(* IEC 61131-3 sources: daoli-st-library/DL_MathData (part 10) *)

(* ---- FC_DL_CharIsAlnum.st ---- *)
(*==============================================================================
 * 组件名称 : FC_DL_CharIsAlnum ｜ 子库 : DL_MathData ｜ v1.0.0 ｜ 2026-11-23
 * 平台     : CODESYS 3.5 / TwinCAT 3 / InoProShop / Machine Expert（纯 IEC，无厂商库）
 * 功能简介 : 判定 STRING(1) 单字符是否为字母或数字（'0'..'9' / 'A'..'Z' /
 *            'a'..'z'），直接以字符（ASCII 序）比较实现，不用库函数。
 * 契约     : 返回 TRUE = 字母或数字；输入 sChar 单字符，空串恒 FALSE；
 *            纯函数无状态、同输入同输出。
 * 开源溯源 : 来源 fisothemes/TwinCAT-Dynamic-String-Kit
 *            https://github.com/fisothemes/TwinCAT-Dynamic-String-Kit / MIT
 *            借鉴点：字符分类谓词语义，实现为本库 clean-room 重写。
 * 依赖     : 无 DL_ 内部依赖（本批自足实现）
 * 红线自检 : R1 零全局 R2 零%I/%Q R3 纯IEC R4 空串防御（区间外恒 FALSE）
 *            R5 双语注释 R6 N/A（无状态机） R7 N/A（无定时器实例）
 * 修订历史 : 2026-11-23 R78-B1 字符分类族模板派生首版
 *============================================================================*)
FUNCTION FC_DL_CharIsAlnum : BOOL
VAR_INPUT
    sChar : STRING(1);      // 待判定单字符（空串恒 FALSE） / Single character to test (empty = FALSE)
END_VAR
IF (sChar >= '0') AND (sChar <= '9') THEN
    FC_DL_CharIsAlnum := TRUE;      // 数字字符命中 / Digit hit
ELSIF ((sChar >= 'A') AND (sChar <= 'Z')) OR ((sChar >= 'a') AND (sChar <= 'z')) THEN
    FC_DL_CharIsAlnum := TRUE;      // 字母字符命中 / Letter hit
ELSE
    FC_DL_CharIsAlnum := FALSE;     // 空串或其他字符 / Empty string or other character
END_IF
END_FUNCTION

(* ---- FC_DL_CharIsAlpha.st ---- *)
(*==============================================================================
 * 组件名称 : FC_DL_CharIsAlpha ｜ 子库 : DL_MathData ｜ v1.0.0 ｜ 2026-11-23
 * 平台     : CODESYS 3.5 / TwinCAT 3 / InoProShop / Machine Expert（纯 IEC，无厂商库）
 * 功能简介 : 判定 STRING(1) 单字符是否为英文字母 'A'..'Z' 或 'a'..'z'，
 *            直接以字符（ASCII 序）比较实现，不调用任何字符分类库函数。
 * 契约     : 返回 TRUE = 英文字母；输入 sChar 单字符，空串按非字母处理；
 *            纯函数无状态、同输入同输出。
 * 开源溯源 : 来源 fisothemes/TwinCAT-Dynamic-String-Kit
 *            https://github.com/fisothemes/TwinCAT-Dynamic-String-Kit / MIT
 *            借鉴点：字符分类谓词语义，实现为本库 clean-room 重写。
 * 依赖     : 无 DL_ 内部依赖（本批自足实现）
 * 红线自检 : R1 零全局 R2 零%I/%Q R3 纯IEC R4 空串防御（区间外恒 FALSE）
 *            R5 双语注释 R6 N/A（无状态机） R7 N/A（无定时器实例）
 * 修订历史 : 2026-11-23 R78-B1 字符分类族模板派生首版
 *============================================================================*)
FUNCTION FC_DL_CharIsAlpha : BOOL
VAR_INPUT
    sChar : STRING(1);      // 待判定单字符（空串按非字母） / Single character to test (empty = not alpha)
END_VAR
IF ((sChar >= 'A') AND (sChar <= 'Z')) OR ((sChar >= 'a') AND (sChar <= 'z')) THEN
    FC_DL_CharIsAlpha := TRUE;      // 命中大小写字母区间 / Within letter ranges A-Z or a-z
ELSE
    FC_DL_CharIsAlpha := FALSE;     // 空串或非字母字符 / Empty string or non-letter
END_IF
END_FUNCTION

(* ---- FC_DL_CharIsDigit.st ---- *)
(*==============================================================================
 * 组件名称 : FC_DL_CharIsDigit ｜ 子库 : DL_MathData ｜ v1.0.0 ｜ 2026-11-23
 * 平台     : CODESYS 3.5 / TwinCAT 3 / InoProShop / Machine Expert（纯 IEC，无厂商库）
 * 功能简介 : 判定 STRING(1) 单字符是否为十进制数字字符 '0'..'9'，
 *            直接以字符（ASCII 序）比较实现，不调用任何字符分类库函数。
 * 契约     : 返回 TRUE = 数字字符；输入 sChar 单字符，空串按非数字处理；
 *            纯函数无状态、同输入同输出。
 * 开源溯源 : 来源 fisothemes/TwinCAT-Dynamic-String-Kit
 *            https://github.com/fisothemes/TwinCAT-Dynamic-String-Kit / MIT
 *            借鉴点：字符分类谓词语义，实现为本库 clean-room 重写。
 * 依赖     : 无 DL_ 内部依赖（本批自足实现）
 * 红线自检 : R1 零全局 R2 零%I/%Q R3 纯IEC R4 空串防御（区间外恒 FALSE）
 *            R5 双语注释 R6 N/A（无状态机） R7 N/A（无定时器实例）
 * 修订历史 : 2026-11-23 R78-B1 字符分类族模板派生首版
 *============================================================================*)
FUNCTION FC_DL_CharIsDigit : BOOL
VAR_INPUT
    sChar : STRING(1);      // 待判定单字符（空串按非数字） / Single character to test (empty = not a digit)
END_VAR
IF (sChar >= '0') AND (sChar <= '9') THEN
    FC_DL_CharIsDigit := TRUE;      // 命中 '0'..'9' 区间 / Within digit range '0'..'9'
ELSE
    FC_DL_CharIsDigit := FALSE;     // 空串或非数字字符 / Empty string or non-digit
END_IF
END_FUNCTION

(* ---- FC_DL_CharIsHexDigit.st ---- *)
(*==============================================================================
 * 组件名称 : FC_DL_CharIsHexDigit ｜ 子库 : DL_MathData ｜ v1.0.0 ｜ 2026-11-23
 * 平台     : CODESYS 3.5 / TwinCAT 3 / InoProShop / Machine Expert（纯 IEC，无厂商库）
 * 功能简介 : 判定 STRING(1) 单字符是否为十六进制位（'0'..'9' / 'A'..'F' /
 *            'a'..'f'），直接以字符（ASCII 序）比较实现，不用库函数。
 * 契约     : 返回 TRUE = 十六进制位；输入 sChar 单字符，空串恒 FALSE；
 *            纯函数无状态、同输入同输出。
 * 开源溯源 : 来源 fisothemes/TwinCAT-Dynamic-String-Kit
 *            https://github.com/fisothemes/TwinCAT-Dynamic-String-Kit / MIT
 *            借鉴点：字符分类谓词语义，实现为本库 clean-room 重写。
 * 依赖     : 无 DL_ 内部依赖（本批自足实现）
 * 红线自检 : R1 零全局 R2 零%I/%Q R3 纯IEC R4 空串防御（恒 FALSE）
 *            R5 双语注释 R6 N/A（无状态机） R7 N/A（无定时器实例）
 * 修订历史 : 2026-11-23 R78-B1 字符分类族模板派生首版
 *============================================================================*)
FUNCTION FC_DL_CharIsHexDigit : BOOL
VAR_INPUT
    sChar : STRING(1);      // 待判定单字符（空串恒 FALSE） / Single character to test (empty = FALSE)
END_VAR
IF (sChar >= '0') AND (sChar <= '9') THEN
    FC_DL_CharIsHexDigit := TRUE;       // 数字位命中 / Decimal digit hit
ELSIF (sChar >= 'A') AND (sChar <= 'F') THEN
    FC_DL_CharIsHexDigit := TRUE;       // 大写十六进制位命中 / Uppercase hex letter hit
ELSIF (sChar >= 'a') AND (sChar <= 'f') THEN
    FC_DL_CharIsHexDigit := TRUE;       // 小写十六进制位命中 / Lowercase hex letter hit
ELSE
    FC_DL_CharIsHexDigit := FALSE;      // 空串或其他字符 / Empty string or other character
END_IF
END_FUNCTION

(* ---- FC_DL_CharIsLower.st ---- *)
(*==============================================================================
 * 组件名称 : FC_DL_CharIsLower ｜ 子库 : DL_MathData ｜ v1.0.0 ｜ 2026-11-23
 * 平台     : CODESYS 3.5 / TwinCAT 3 / InoProShop / Machine Expert（纯 IEC，无厂商库）
 * 功能简介 : 判定 STRING(1) 单字符是否为小写英文字母 'a'..'z'，
 *            直接以字符（ASCII 序）比较实现，不调用任何字符分类库函数。
 * 契约     : 返回 TRUE = 小写字母；输入 sChar 单字符，空串恒 FALSE；
 *            纯函数无状态、同输入同输出。
 * 开源溯源 : 来源 fisothemes/TwinCAT-Dynamic-String-Kit
 *            https://github.com/fisothemes/TwinCAT-Dynamic-String-Kit / MIT
 *            借鉴点：字符分类谓词语义，实现为本库 clean-room 重写。
 * 依赖     : 无 DL_ 内部依赖（本批自足实现）
 * 红线自检 : R1 零全局 R2 零%I/%Q R3 纯IEC R4 空串防御（区间外恒 FALSE）
 *            R5 双语注释 R6 N/A（无状态机） R7 N/A（无定时器实例）
 * 修订历史 : 2026-11-23 R78-B1 字符分类族模板派生首版
 *============================================================================*)
FUNCTION FC_DL_CharIsLower : BOOL
VAR_INPUT
    sChar : STRING(1);      // 待判定单字符（空串恒 FALSE） / Single character to test (empty = FALSE)
END_VAR
IF (sChar >= 'a') AND (sChar <= 'z') THEN
    FC_DL_CharIsLower := TRUE;      // 命中 'a'..'z' 区间 / Within lowercase range 'a'..'z'
ELSE
    FC_DL_CharIsLower := FALSE;     // 空串或非小写字母 / Empty string or not lowercase
END_IF
END_FUNCTION

(* ---- FC_DL_CharIsSpace.st ---- *)
(*==============================================================================
 * 组件名称 : FC_DL_CharIsSpace ｜ 子库 : DL_MathData ｜ v1.0.0 ｜ 2026-11-23
 * 平台     : CODESYS 3.5 / TwinCAT 3 / InoProShop / Machine Expert（纯 IEC，无厂商库）
 * 功能简介 : 判定 STRING(1) 单字符是否为空白字符（空格 16#20 或水平制表符
 *            Tab 16#09），Tab 用 IEC 标准字符串转义 '$T' 表示，不用库函数。
 * 契约     : 返回 TRUE = 空格或 Tab；输入 sChar 单字符，空串恒 FALSE；
 *            纯函数无状态、同输入同输出。
 * 开源溯源 : 来源 fisothemes/TwinCAT-Dynamic-String-Kit
 *            https://github.com/fisothemes/TwinCAT-Dynamic-String-Kit / MIT
 *            借鉴点：字符分类谓词语义，实现为本库 clean-room 重写。
 * 依赖     : 无 DL_ 内部依赖（本批自足实现）
 * 红线自检 : R1 零全局 R2 零%I/%Q R3 纯IEC（'$T' 为 IEC 标准转义）
 *            R4 空串防御（恒 FALSE） R5 双语注释 R6 N/A（无状态机） R7 N/A（无定时器实例）
 * 修订历史 : 2026-11-23 R78-B1 字符分类族模板派生首版
 *============================================================================*)
FUNCTION FC_DL_CharIsSpace : BOOL
VAR_INPUT
    sChar : STRING(1);      // 待判定单字符（空串恒 FALSE） / Single character to test (empty = FALSE)
END_VAR
IF (sChar = ' ') OR (sChar = '$T') THEN
    FC_DL_CharIsSpace := TRUE;      // 空格或 Tab 命中 / Space or tab hit
ELSE
    FC_DL_CharIsSpace := FALSE;     // 空串或其他字符 / Empty string or other character
END_IF
END_FUNCTION

(* ---- FC_DL_CharIsUpper.st ---- *)
(*==============================================================================
 * 组件名称 : FC_DL_CharIsUpper ｜ 子库 : DL_MathData ｜ v1.0.0 ｜ 2026-11-23
 * 平台     : CODESYS 3.5 / TwinCAT 3 / InoProShop / Machine Expert（纯 IEC，无厂商库）
 * 功能简介 : 判定 STRING(1) 单字符是否为大写英文字母 'A'..'Z'，
 *            直接以字符（ASCII 序）比较实现，不调用任何字符分类库函数。
 * 契约     : 返回 TRUE = 大写字母；输入 sChar 单字符，空串恒 FALSE；
 *            纯函数无状态、同输入同输出。
 * 开源溯源 : 来源 fisothemes/TwinCAT-Dynamic-String-Kit
 *            https://github.com/fisothemes/TwinCAT-Dynamic-String-Kit / MIT
 *            借鉴点：字符分类谓词语义，实现为本库 clean-room 重写。
 * 依赖     : 无 DL_ 内部依赖（本批自足实现）
 * 红线自检 : R1 零全局 R2 零%I/%Q R3 纯IEC R4 空串防御（区间外恒 FALSE）
 *            R5 双语注释 R6 N/A（无状态机） R7 N/A（无定时器实例）
 * 修订历史 : 2026-11-23 R78-B1 字符分类族模板派生首版
 *============================================================================*)
FUNCTION FC_DL_CharIsUpper : BOOL
VAR_INPUT
    sChar : STRING(1);      // 待判定单字符（空串恒 FALSE） / Single character to test (empty = FALSE)
END_VAR
IF (sChar >= 'A') AND (sChar <= 'Z') THEN
    FC_DL_CharIsUpper := TRUE;      // 命中 'A'..'Z' 区间 / Within uppercase range 'A'..'Z'
ELSE
    FC_DL_CharIsUpper := FALSE;     // 空串或非大写字母 / Empty string or not uppercase
END_IF
END_FUNCTION

(* ---- FC_DL_CharToUpper.st ---- *)
(*==============================================================================
 * 组件名称 : FC_DL_CharToUpper ｜ 子库 : DL_MathData ｜ v1.0.0 ｜ 2026-11-23
 * 平台     : CODESYS 3.5 / TwinCAT 3 / InoProShop / Machine Expert（纯 IEC，无厂商库）
 * 功能简介 : 小写英文字母转大写（'a'..'z' → 'A'..'Z'），其余字符原样返回。
 *            无字符算术库函数可用，故以 26 项等值映射（每行两项）实现，
 *            语义与 ASCII 减 32 完全一致。
 * 契约     : 返回转换后的单字符；输入 sChar 单字符；空串原样返回；
 *            纯函数无状态、同输入同输出。
 * 开源溯源 : 来源 fisothemes/TwinCAT-Dynamic-String-Kit
 *            https://github.com/fisothemes/TwinCAT-Dynamic-String-Kit / MIT
 *            借鉴点：字符分类/变换谓词语义，实现为本库 clean-room 重写。
 * 依赖     : 无 DL_ 内部依赖（本批自足实现）
 * 红线自检 : R1 零全局 R2 零%I/%Q R3 纯IEC R4 空串原样返回无越界
 *            R5 双语注释 R6 N/A（无状态机） R7 N/A（无定时器实例）
 * 修订历史 : 2026-11-23 R78-B1 字符分类族模板派生首版
 *============================================================================*)
FUNCTION FC_DL_CharToUpper : STRING(1)
VAR_INPUT
    sChar : STRING(1);      // 待转换单字符 / Single character to convert
END_VAR
IF sChar = 'a' THEN FC_DL_CharToUpper := 'A'; ELSIF sChar = 'b' THEN FC_DL_CharToUpper := 'B';        // a→A b→B a/b to upper
ELSIF sChar = 'c' THEN FC_DL_CharToUpper := 'C'; ELSIF sChar = 'd' THEN FC_DL_CharToUpper := 'D';     // c→C d→D c/d to upper
ELSIF sChar = 'e' THEN FC_DL_CharToUpper := 'E'; ELSIF sChar = 'f' THEN FC_DL_CharToUpper := 'F';     // e→E f→F e/f to upper
ELSIF sChar = 'g' THEN FC_DL_CharToUpper := 'G'; ELSIF sChar = 'h' THEN FC_DL_CharToUpper := 'H';     // g→G h→H g/h to upper
ELSIF sChar = 'i' THEN FC_DL_CharToUpper := 'I'; ELSIF sChar = 'j' THEN FC_DL_CharToUpper := 'J';     // i→I j→J i/j to upper
ELSIF sChar = 'k' THEN FC_DL_CharToUpper := 'K'; ELSIF sChar = 'l' THEN FC_DL_CharToUpper := 'L';     // k→K l→L k/l to upper
ELSIF sChar = 'm' THEN FC_DL_CharToUpper := 'M'; ELSIF sChar = 'n' THEN FC_DL_CharToUpper := 'N';     // m→M n→N m/n to upper
ELSIF sChar = 'o' THEN FC_DL_CharToUpper := 'O'; ELSIF sChar = 'p' THEN FC_DL_CharToUpper := 'P';     // o→O p→P o/p to upper
ELSIF sChar = 'q' THEN FC_DL_CharToUpper := 'Q'; ELSIF sChar = 'r' THEN FC_DL_CharToUpper := 'R';     // q→Q r→R q/r to upper
ELSIF sChar = 's' THEN FC_DL_CharToUpper := 'S'; ELSIF sChar = 't' THEN FC_DL_CharToUpper := 'T';     // s→S t→T s/t to upper
ELSIF sChar = 'u' THEN FC_DL_CharToUpper := 'U'; ELSIF sChar = 'v' THEN FC_DL_CharToUpper := 'V';     // u→U v→V u/v to upper
ELSIF sChar = 'w' THEN FC_DL_CharToUpper := 'W'; ELSIF sChar = 'x' THEN FC_DL_CharToUpper := 'X';     // w→W x→X w/x to upper
ELSIF sChar = 'y' THEN FC_DL_CharToUpper := 'Y'; ELSIF sChar = 'z' THEN FC_DL_CharToUpper := 'Z';     // y→Y z→Z y/z to upper
ELSE
    FC_DL_CharToUpper := sChar;     // 非小写字母（含空串/大写/符号）原样返回 / Non-lowercase returned unchanged
END_IF
END_FUNCTION

(* ---- FC_DL_ChecksumLwordSum.st ---- *)
(*
  Name        : FC_DL_ChecksumLwordSum
  Category    : DL_MathData
  Version     : 1.0.0
  Purpose     : 64 位字累加和校验：LWORD 数组按模 2^64 回卷累加（高低半字条件进位，禁取模），与预置校验值位等比对出结论；/ 64-bit word checksum: modulo-2^64 wrapping accumulate of an LWORD array via conditional halfword carry (no modulo), compared bit-equal against a preset check value
  溯源        : 借 lgf-datahandling 的分类/参数域组织，clean-room 实现
  Boundary    : ① 空数组（计数 0）→ 返回 FALSE 哨兵，不返回 0 当有效和；
                ② 回卷累加用条件进位法（低半字加后回卷即进位），全程禁取模运算；
                ③ 数组长度上限常量守卫 + 计数域闸（负数/超容拒绝），遍历用 FOR 有界循环防死循环；
                ④ 预置校验值比对为整数位等（无浮点判等）；
                ⑤ 高半字加法回卷即模 2^64 语义（溢出进位出界自然丢弃）；
                ⑥ 本件为纯函数：无状态、无实例保持量、零外部全局、零物理地址。
*)
FUNCTION FC_DL_ChecksumLwordSum : BOOL
VAR_INPUT
    aData   : ARRAY[1..256] OF LWORD;        (* 待校验数据数组（有效区 1..nCount）[-] / Data array to checksum *)
    nCount  : INT := 0;                      (* 有效元素计数，域 0..256 [-] / Valid element count *)
    qwExpect: LWORD := LWORD#0;              (* 预置校验值（位等比对目标）[-] / Preset expected checksum *)
END_VAR
VAR_OUTPUT
    qwSum   : LWORD;                         (* 累加和出口（空数组时为 0 且返回 FALSE）[-] / Accumulated sum outlet *)
    bMatch  : BOOL;                          (* 比对结论：累加和与预置值位等 [-] / Match verdict, bit-equal *)
END_VAR
VAR
    _nCnt   : INT;                           (* 钳位后生效元素计数 [个] / Clamped element count *)
    _i      : INT;                           (* 遍历游标 [个] / Loop cursor *)
    _sLo    : DWORD;                         (* 累加和低半字 [-] / Sum low halfword *)
    _sHi    : DWORD;                         (* 累加和高半字 [-] / Sum high halfword *)
    _tLo    : DWORD;                         (* 低半字加法暂存（回卷检测）[-] / Low half add staging *)
    _tHi    : DWORD;                         (* 高半字加法暂存（回卷丢弃）[-] / High half add staging *)
    _eLo    : DWORD;                         (* 当前元素低半字 [-] / Element low half *)
    _eHi    : DWORD;                         (* 当前元素高半字 [-] / Element high half *)
    _cIn    : DWORD;                         (* 低半字回卷进位（0/1）[-] / Carry from low wrap *)
END_VAR
VAR CONSTANT
    DL_CKS_NMAX  : INT   := 256;             (* 数组容量上限常量守卫 [个] / Array capacity guard *)
    DL_CKS_MASKL : LWORD := LWORD#16#FFFFFFFF;   (* 低 32 位掩码常量 [-] / Low 32-bit mask *)
END_VAR

(* —— 段 1：出口与累加器预清（空数组哨兵前置，R107） —— *)
qwSum  := LWORD#0;                                       (* 累加和出口预清（哨兵零） / Sum outlet preset *)
bMatch := FALSE;                                         (* 比对结论预清 / Match preset *)
_sLo := DWORD#0;                                         (* 低半字累加清零 / Low half clear *)
_sHi := DWORD#0;                                         (* 高半字累加清零 / High half clear *)

(* —— 段 2：计数域闸 + 容量守卫（边界③） —— *)
_nCnt := nCount;                                         (* 生效计数初值 / Effective count init *)
IF (nCount < 0) OR (nCount > DL_CKS_NMAX) THEN
    FC_DL_ChecksumLwordSum := FALSE;                     (* 计数越域：哨兵拒绝（不出有效和） / Count out of domain, sentinel reject *)
    RETURN;                                              (* 提前返回（无状态残留） / Early return *)
END_IF
IF _nCnt = 0 THEN
    FC_DL_ChecksumLwordSum := FALSE;                     (* 空数组：哨兵拒绝，不返回 0 当有效和（边界①） / Empty array, sentinel reject *)
    RETURN;                                              (* 提前返回 / Early return *)
END_IF

(* —— 段 3：条件进位回卷累加（禁取模，边界②⑤；FOR 有界防死循环） —— *)
FOR _i := 1 TO _nCnt DO
    _eLo := LWORD_TO_DWORD(aData[_i] AND DL_CKS_MASKL);  (* 取元素低半字（掩码常量） / Element low half *)
    _eHi := LWORD_TO_DWORD(SHR(aData[_i], 32));          (* 取元素高半字（移 32 位常量） / Element high half *)
    _tLo := _sLo + _eLo;                                 (* 低半字相加 / Low half add *)
    IF _tLo < _sLo THEN
        _cIn := DWORD#1;                                 (* 回卷即进位（条件进位法） / Wrap implies carry *)
    ELSE
        _cIn := DWORD#0;                                 (* 无回卷无进位 / No carry *)
    END_IF
    _sLo := _tLo;                                        (* 低半字推进 / Low half advance *)
    _tHi := _sHi + _eHi + _cIn;                          (* 高半字带进位相加 / High half add with carry *)
    _sHi := _tHi;                                        (* 高半字回卷进位出界自然丢弃（模 2^64 语义） / High wrap discard *)
END_FOR

(* —— 段 4：出口组装 + 位等比对（边界④，整数无浮点） —— *)
qwSum  := SHL(DWORD_TO_LWORD(_sHi), 32) OR DWORD_TO_LWORD(_sLo);   (* 半字合成 64 位和 / Assemble 64-bit sum *)
bMatch := (qwSum = qwExpect);                            (* 位等比对（整数直比） / Bit-equal compare *)
FC_DL_ChecksumLwordSum := TRUE;                          (* 有效和结论 / Valid sum verdict *)
END_FUNCTION

(* ---- FC_DL_ChecksumSum64.st ---- *)
// =====================================================================
// FC_DL_ChecksumSum64.st
// LWORD 数组 64 位累加和校验（纯函数, 模 2^64 自然回绕求和 + 越界守卫）
// 64-bit LWORD array additive checksum, pure function
// 所属子库: DL_MathData    版本: v1.0.0    兼容: CODESYS V3.5+ / TwinCAT 3 / 汇川 InoProShop
// 码位: 16#0001_048A ~ 16#0001_048D (本件独占 4 槽, FC 纯函数分型, 勿复用)
// 溯源: IEC 61131-3 标准语义的道莅防御性实现
//       来源组标签: checksum, data-integrity, pure-function, lword
// 修改记录: R30 初版 (ROUND_PLAN_R30 序 19)
// 语义声明: 模 2^64 累加和由 LWORD 无符号加法自然回绕实现, 禁用取余运算;
//           与 FC_DL_ChecksumSum8 构成 8/64 位宽两件, 位宽变体不再扩充;
//           错误出口约定与 FC_DL_ChecksumSum8 现行 uErrorId 出口一致;
//           纯函数无内部状态, 码为返回拍瞬时值, 无锁存面
// =====================================================================
FUNCTION FC_DL_ChecksumSum64 : LWORD   // 返回累加和, 异常路径返回哨兵零值 / Returns sum, sentinel zero on fault
VAR_INPUT
    aData  : ARRAY[*] OF LWORD;     // 被校验数组（开数组, 实测边界）/ Data array, open bounds
    uCount : USINT;                 // 参与求和的元素个数 1~255 / Element count
END_VAR
VAR_OUTPUT
    uErrorId : UDINT;               // 错误码, 见码表 / Error code, see table
END_VAR
VAR
    uCap   : DINT := 0;             // 数组实测元素容量 / Measured array capacity
    uNum   : DINT := 0;             // 钳位后的求和个数 / Effective count
    iIdx   : DINT := 0;             // 循环下标 / Loop index
    iElem  : DINT := 0;             // 数组元素下标 / Element index
    lwSum  : LWORD := LWORD#0;      // 累加和 / Accumulated sum
    lwPrev : LWORD := LWORD#0;      // 上拍和快照（回绕检测）/ Previous sum for wrap detect
    xWrap  : BOOL := FALSE;         // 自然回绕发生标记 / Wraparound occurred flag
END_VAR

// ---------------------------------------------------------------------
// 代码位表（本件独占, 勿复用）:
//   16#0001_048A 信息 累加和计算完成（含自然回绕路径）
//   16#0001_048B 信息 空输入（计数为 0, 返回哨兵零值）
//   16#0001_048C 故障 计数越界（大于数组实测容量, 强制退出, 返回零值）,
//                纯函数无锁存面, 修正入参重新调用即解除
//   16#0001_048D 信息 求和自然回绕发生（本拍回绕旁证, 供数据链路诊断）
// ---------------------------------------------------------------------

// ---- 缺省返回哨兵零值 / Default sentinel zero ----
FC_DL_ChecksumSum64 := LWORD#0;

// ---- 容量实测（开数组边界实测, 不假设下标起点）/ Measured capacity ----
IF UPPER_BOUND(aData, 1) >= LOWER_BOUND(aData, 1) THEN
    uCap := (UPPER_BOUND(aData, 1) - LOWER_BOUND(aData, 1)) + 1;    // 元素个数 / Element count
END_IF

// ---- 空输入: 计数为 0, 返回哨兵零 + 信息码 / Empty input ----
IF uCount = 0 THEN
    uErrorId := 16#0001_048B;       // 空输入码 / Empty input code
    RETURN;                         // 返回零值 / Return zero
END_IF

// ---- 计数越界守护: 强制退出 / Count overrun guard: force exit ----
uNum := USINT_TO_DINT(uCount);
IF uNum > uCap THEN
    uErrorId := 16#0001_048C;       // 越界故障码 / Overrun fault code
    RETURN;                         // 强制退出返回零 / Force exit with zero
END_IF

// ---- 模 2^64 累加（LWORD 自然回绕, 禁用取余）/ Modulo sum by natural wrap ----
lwSum := LWORD#0;                   // 和清零 / Clear sum
xWrap := FALSE;                     // 回绕标记复位 / Reset wrap flag
FOR iIdx := 1 TO uNum DO
    iElem := LOWER_BOUND(aData, 1) + (iIdx - 1);    // 实测下标映射 / Measured index mapping
    lwPrev := lwSum;                // 上拍和快照 / Snapshot previous sum
    lwSum := lwSum + aData[iElem];  // 累加（无符号自然回绕）/ Accumulate with natural wrap
    IF lwSum < lwPrev THEN
        xWrap := TRUE;              // 无符号回绕旁证 / Unsigned wrap occurred
    END_IF
END_FOR

FC_DL_ChecksumSum64 := lwSum;       // 返回累加和 / Return sum
IF xWrap THEN
    uErrorId := 16#0001_048D;       // 回绕旁证码 / Wrap hint code
ELSE
    uErrorId := 16#0001_048A;       // 完成码 / Done code
END_IF

END_FUNCTION

(* ---- FC_DL_ChecksumSum8.st ---- *)
(*
    组件名称 : FC_DL_ChecksumSum8
    所属子库 : DL_MathData
    当前版本 : 1.0.0
    兼 容 性 : CODESYS V3.5+ / TwinCAT 3 / 汇川 InoProShop；仅依赖 Standard.library
    功能描述 : 8 位累加和校验，覆盖 DL/T 645、水表/电表自定义帧这类「不用 CRC、只用累加和」的协议形态。
              取舍 ①：用 DINT 累加而不是 BYTE 累加 —— 255 × 256 在 BYTE 域必然回绕，回绕本身虽等价于 MOD 256，
              但一旦有人在中间插入一步「判和是否超限」的诊断，回绕后的和就已经撒谎；升位累加、末了一次取模，
              中间量始终可观测。
              取舍 ②：补码模式的结果 0 必须显式判 —— 累加和 0 的补码在数学上仍是 0（不是 256），
              若写成 256 − 0 会溢出成 256 再被截成 0，看着对但依赖隐式回绕；而且「校验字节为 0」在部分协议里
              表示「本帧无校验」，这条歧义必须发信息码让上位机知情。
              取舍 ③：帧长超上限拒绝而不截断 —— 同 CRC 件口径，截断后的累加和格式合法但必然校验失败。
              取舍 ④：本件不做 LWORD 累加变体 —— 64 位累加和没有任何公开协议用例，属过度设计，
              8 位才是实际协议形态；该判断已在本轮规格留档。
    开源溯源 : T2-1 LGF Data Handling 子族（「校验族尚余累加和待挖」）；算法为公开经典，零查表、；本件为道莅 clean-room 防御性实现（仅借 LGF 分类事实/参数域/行为定义，零代码行与符号名复制）。
              零代码行复制，码位与分级 100% 自有。
    本文件内含 : FUNCTION FC_DL_ChecksumSum8（单 POU，无配套类型）
    依 赖 : 无 DL_ 内部依赖；Standard.library: 无
    红线自检 : R1 ✓ 零全局变量与外部变量 ｜ R2 ✓ 零物理 IO 地址
              R3 ✓ 纯 IEC 61131-3 ｜ R4 ✓ 帧长闸 + 空帧短路 + 补码零特例 + 累加升位防回绕 + 取模前操作数非负
              R5 ✓ 全变量中英双语同行注释 ｜ R6 N/A 纯函数无顺序状态机，无 CASE 可写
              R7 N/A 无定时器、无沿检测实例 ｜ R8 ✓ 取模基数与缓冲上限常量化
    错误码   : 16#0001_0446 [信息级] 补码模式下结果为 0 的特例（部分协议以 0 表示无校验），bValid = TRUE
               16#0001_0447 [信息级] 空帧，返回 0，bValid = TRUE
               16#0001_0387 [故障级] 帧长超 DL_SUM_BUF_MAX，拒绝计算，返回 0，bValid = FALSE
               16#0001_0388 [故障级] 预留禁用（不得挪用）
               16#0001_0389 [故障级] 预留禁用（不得挪用）
    码位总账 : 16#0001_0446 用 / 16#0001_0447 用 ｜ 16#0001_0387 用 / 16#0001_0388 预留 / 16#0001_0389 预留
    遗留假设 : ① 累加上界推导：最大 255 × 255 + 255 级余量远小于 DINT 上界，中间量不会溢出；
              该推导依赖「nLen ≤ 255 由闸门保证」，若上限常量被改大须重新核算（已在头注释留痕）。
              ② 无内建转换链依赖，编译门槛未见风险。
    修订历史 :
        2026-11-16  v1.0.0  首版，R21 批次 2 入库
*)
FUNCTION FC_DL_ChecksumSum8 : BYTE
VAR_INPUT
    nLen            : UINT;   // 待累加字节数，0~DL_SUM_BUF_MAX，0 = 空帧 [字节] / number of bytes, zero means an empty frame [byte]
    bTwosComplement : BOOL := FALSE;   // TRUE 输出累加和的二进制补码（DL/T 645 口径）/ TRUE returns the two's complement, the DL/T 645 convention
END_VAR
VAR_IN_OUT
    afData          : ARRAY[0..DL_SUM_BUF_MAX] OF BYTE;   // 待累加字节数组，仅前 nLen 个有效 [字节] / data buffer, only the first nLen bytes are used [byte]
END_VAR
VAR_OUTPUT
    eErr            : UDINT;  // 错误码，0=正常；16#0001_04XX 信息级 / 16#0001_03XX 故障级 / error id, 0=ok
    bError          : BOOL;   // 故障级标志，eErr 落 16#0001_03XX 时为 TRUE / fault flag, TRUE on fault-level eErr
    bValid          : BOOL;   // 返回值是否可用 / result usable flag
END_VAR
VAR
    nSum            : DINT;   // 升位累加器，恒非负 [无量纲] / widened accumulator, always non-negative [dimensionless]
    nModRes         : DINT;   // 累加和对 256 取模后的低 8 位值 [无量纲] / low byte value after the modulo [dimensionless]
    uIdx            : UINT;   // 字节游标 [字节] / byte cursor [byte]
    uRet            : BYTE;   // 校验字节结果 [字节] / checksum byte result [byte]
END_VAR
VAR CONSTANT
    DL_SUM_BUF_MAX  : UINT := 255;     // 单帧字节数上限 [字节] / frame length upper bound [byte]
    DL_BYTE_MOD     : DINT := 256;     // 8 位容器的取模基数 [无量纲] / modulus of the byte container [dimensionless]
    DL_DINT_ZERO    : DINT := 0;       // 零哨兵 [无量纲] / zero sentinel [dimensionless]
    DL_SUM_LEN_NONE : UINT := 0;       // 空帧长度哨兵，减法前必判 [字节] / empty frame sentinel [byte]
    DL_BYTE_ZERO    : BYTE := 16#00;   // 字节零哨兵 [字节] / byte zero sentinel [byte]
    DL_ERR_NONE     : UDINT := 16#0000_0000;   // 无故障 / no error
END_VAR

// 段 1｜返回值与错误状态预置 / segment 1, preset the return value and the error state
FC_DL_ChecksumSum8 := DL_BYTE_ZERO;   // 故障缺省返回 0 / fault default returns zero
eErr   := DL_ERR_NONE;                // 预置无错误 / preset no error
bError := FALSE;                      // 预置无故障 / preset no fault
bValid := FALSE;                      // 预置结果不可用 / preset unusable
nSum   := DL_DINT_ZERO;               // 累加器清零 / clear the accumulator

// 段 2｜帧长闸：超上限拒绝，绝不截断 / segment 2, length gate, refuse instead of truncating
IF nLen > DL_SUM_BUF_MAX THEN
    eErr   := 16#0001_0387;           // 帧长超上限（故障级）/ frame too long, fault level
    bError := TRUE;                   // 置故障标志 / raise the fault flag
    RETURN;                           // 返回 0，bValid 保持 FALSE / return zero, bValid stays FALSE
END_IF

// 段 3｜空帧短路：长度 0 时 nLen − 1 会回绕成 65535，必须先判零 / segment 3, empty frame short circuit before any subtraction
IF nLen = DL_SUM_LEN_NONE THEN
    FC_DL_ChecksumSum8 := DL_BYTE_ZERO;   // 空帧累加和为 0 / an empty frame sums to zero
    eErr   := 16#0001_0447;               // 空帧（信息级，不置 bError）/ empty frame, info level
    bValid := TRUE;                       // 空帧是协议合法输入 / an empty frame is a legal protocol input
    RETURN;                               // 提前出口，绝不进循环 / early exit, never enter the loop
END_IF

// 段 4｜升位累加：nLen 已保证 ≥ 1 / segment 4, widened accumulation, nLen is at least one
FOR uIdx := 0 TO nLen - 1 DO
    nSum := nSum + BYTE_TO_DINT(afData[uIdx]);   // 升到 DINT 累加，中间量始终可观测 / widen to DINT so the intermediate stays observable
END_FOR

// 段 5｜取模与补码：nSum 恒非负，MOD 安全 / segment 5, modulo and two's complement, the operand is never negative
nModRes := nSum MOD DL_BYTE_MOD;      // 低 8 位值，0~255 / the low byte, 0..255
IF bTwosComplement THEN
    IF nModRes = DL_DINT_ZERO THEN
        uRet := DL_BYTE_ZERO;         // 零的补码仍是零，显式判，不依赖 256 − 0 的回绕 / zero complements to zero, tested explicitly
        eErr := 16#0001_0446;         // 补码结果为零的特例（信息级）/ two's complement result is zero, info level
    ELSE
        uRet := DINT_TO_BYTE(DL_BYTE_MOD - nModRes);   // 256 − 和，落 1~255 / two hundred and fifty six minus the sum, 1..255
    END_IF
ELSE
    uRet := DINT_TO_BYTE(nModRes);    // 直接取低 8 位 / take the low byte directly
END_IF

// 段 6｜出口 / segment 6, exit
FC_DL_ChecksumSum8 := uRet;           // 输出校验字节 / publish the checksum byte
bValid := TRUE;                       // 结果可用 / the result is usable
END_FUNCTION

(* ---- FC_DL_CircularMeanCalc.st ---- *)
(*
  ==================================================================
  组件名 Component  : FC_DL_CircularMeanCalc
  分类   Category   : DL_MathData
  版本   Version    : 1.0.0
  功能   Purpose    : 角度集的圆均值（Circular Mean）：Σsin/Σcos 合成向量法，
                      输出归一 [0,360) 的平均角。归一采用「条件加减」搬区间
                      （负角加 360 / 满 360 减 360），禁负数取模（MOD 在实数
                      域三平台余数符号不一致）。零向量退化（|R| < 1E-6，各角
                      完全对消）判定失效返回，不做伪输出。
  来源   Source     : t2-1-lgf-measurement（测量族：向量合成求圆均值为公开
                      数学口径，实现零源码复制）
  互引   Cross-ref  : FC_DL_WrapAngleDeg（同族角度归一原子，本件内联了等价
                      [0,360) 搬移逻辑，避免跨件调用改变 FC 返回契约）；
                      FC_DL_AngleDiffWrap（下游做两均值角差用）
  平台   Platform   : 纯 IEC 61131-3 四则 + SIN/COS/SQRT/ATAN2 标准数学函数
                      （三平台 MATH 内建：CODESYS Math.library / TwinCAT
                      TC Math / InoProShop Math）
  依赖   Depends    : 无 DL_ 内部依赖
  设计偏差 Deviation: nCount > 数组实际长度时按数组长度钳位接管（防御性，头注
                      声明，不静默越界；错误码表未为此设码，见码位反证）
  红线   Redline    : R1 零全局/VAR_EXTERNAL/R2 零 %I/%Q/R3 纯 IEC 标准
                      R4 元素级非有限闸 + 除法分母显式闸 + 归一域内安全
                      R5 全变量双语同行注释/R6 纯函数无状态机（CASE 不适用）
                      R7 无定时器与沿检测/R8 容差与循环界全常量化
  错误码 Codes      : 01【失效级】空输入（nCount=0），返回 0，bValid=FALSE
                      02【失效级】任一元素非有限（NaN/±Inf），返回 0
                      03【失效级】零向量退化 |R|<1E-6（各角完全对消），返回 0
  码位反证 Note     : 01/02/03 三码分立依据（R90）：01 无效在输入计数层即可
                      观测、02 无效在元素层、03 无效仅在合成结果层，三者的
                      排查入口不同，不可合并；
                      「nCount 超数组长度钳位」与 01 输出组合不可区分（都按
                      实际长度推进、无独立输出通道），按 R 反证条款不为它设码。
  验收   Acceptance : V1 {10, 350} → 0 ｜ V2 {0, 120, 240} → |R|=0 码 03 ｜
                      V3 空 → 码 01 ｜ V4 含 NaN → 码 02 ｜ V5 单元素 → 自身
  变更   Revision   : 2026-11-22  v1.0.0  R66 首版（编码阶段批 1 序 3）
  ==================================================================
*)
FUNCTION FC_DL_CircularMeanCalc : LREAL
VAR_INPUT
    aAnglesDeg : ARRAY[*] OF LREAL;  // 角度数组 [°] / the angle array [deg]
    nCount     : UDINT;              // 参与计算的角度个数 [个]，超出数组长度按长度钳位 / the count, clamped to the array length
END_VAR
VAR_OUTPUT
    bValid     : BOOL;               // 平均角可用标志 [-] / the mean angle usable flag
    nErrId     : UDINT;              // 错误码，0=正常，01/02/03 见头注 [码] / the error code [code]
END_VAR
VAR
    fxSum      : LREAL;              // Σcos 分量 [无量纲] / the summed cosine component [dimensionless]
    fySum      : LREAL;              // Σsin 分量 [无量纲] / the summed sine component [dimensionless]
    fRad       : LREAL;              // 当前元素弧度 [rad] / the current element in radians [rad]
    fR         : LREAL;              // 合成向量模 [无量纲] / the resultant magnitude [dimensionless]
    fMean      : LREAL;              // 圆均值工作寄存器 [°] / the mean working register [deg]
    uUsed      : UDINT;              // 实际参与个数（钳位后）[个] / the used count after clamping [count]
    uLen       : UDINT;              // 数组实际长度 [个] / the actual array length [count]
    i          : UDINT;              // 循环变量，有界 [索引] / the loop index, bounded [index]
END_VAR
VAR CONSTANT
    CMC_DEG2RAD : LREAL := 0.017453292519943295; // π/180，度转弧度 [rad/°] / pi over 180 [rad per deg]
    CMC_DEG_TURN: LREAL := 360.0;                // 一整圈 [°] / one full turn [deg]
    CMC_R_MIN   : LREAL := 1.0E-6;               // 零向量退化阈值 |R| / the degenerate resultant threshold
    CMC_ERR_NONE : UDINT := 16#0000_0000;        // 无错误 [码] / no error [code]
    CMC_ERR_EMPTY: UDINT := 16#0000_0001;        // 码 01：空输入 / code 01, empty input
    CMC_ERR_NAN  : UDINT := 16#0000_0002;        // 码 02：非有限元素 / code 02, non finite element
    CMC_ERR_ZEROV: UDINT := 16#0000_0003;        // 码 03：零向量退化 / code 03, degenerate zero vector
END_VAR

// 段 1｜输出预置 / segment 1, preset the outputs
FC_DL_CircularMeanCalc := 0.0;  // 失效缺省返回 0 / fault default returns zero
bValid := FALSE;                // 预置不可用 / preset unusable
nErrId := CMC_ERR_NONE;         // 预置无错误 / preset no error
fxSum  := 0.0;                  // 分量累加器清零 / clear the cosine accumulator
fySum  := 0.0;                  // 分量累加器清零 / clear the sine accumulator

// 段 2｜数组长度闸与空闸（结构 RETURN 早退）/ segment 2, array length gate and the empty gate
uLen := UDINT#0;                                        // 预置长度 / preset the length
IF UPPER_BOUND(aAnglesDeg, 1) >= 0 THEN                 // 防御：变长数组上界有效性 / defensive: variable array bound check
    uLen := DINT_TO_UDINT(1 + UPPER_BOUND(aAnglesDeg, 1) - LOWER_BOUND(aAnglesDeg, 1)); // 实际长度（守卫内恒非负）/ the actual length, non negative inside the guard
END_IF
IF nCount = UDINT#0 THEN        // 空输入（码 01）/ empty input, code 01
    nErrId := CMC_ERR_EMPTY;
    RETURN;
END_IF
uUsed := nCount;                                        // 先取原始个数 / take the raw count first
IF uUsed > uLen THEN
    uUsed := uLen;                                      // 超长钳位接管（头注偏差声明）/ clamp to the actual length, documented deviation
END_IF
IF uUsed = UDINT#0 THEN         // 钳位后为空（空数组 + 非零 nCount）→ 仍判空码 / still empty after clamping
    nErrId := CMC_ERR_EMPTY;
    RETURN;
END_IF

// 段 3｜分量累加：元素级非有限闸（码 02）与循环下标闸（uUsed ≤ uLen 已证）
//      segment 3, accumulate components with the per element finite gate and a proven index bound
FOR i := 0 TO UDINT_TO_DINT(uUsed) - 1 DO               // 有界 FOR，上界 uUsed ≤ uLen / bounded loop
    fRad := aAnglesDeg[i] * CMC_DEG2RAD;                // 度转弧度 [rad] / degrees to radians [rad]
    IF (aAnglesDeg[i] <> aAnglesDeg[i]) OR (ABS(aAnglesDeg[i]) > 1.7976931348623157E308) THEN  // 自反判 NaN + 有限域 / reflexive NaN and finiteness
        nErrId := CMC_ERR_NAN;                          // 码 02：非有限元素 / code 02, non finite element
        RETURN;                                         // 结构早退，返回 0 / structural early return
    END_IF
    fxSum := fxSum + COS(fRad);                         // 累加 cos 分量 / accumulate the cosine component
    fySum := fySum + SIN(fRad);                         // 累加 sin 分量 / accumulate the sine component
END_FOR

// 段 4｜零向量退化闸（码 03）：|R| < 1E-6 视为完全对消 / segment 4, the degenerate vector gate
fR := SQRT(fxSum * fxSum + fySum * fySum);              // 合成向量模（被开方数恒非负）/ the resultant magnitude
IF fR < CMC_R_MIN THEN
    nErrId := CMC_ERR_ZEROV;                            // 码 03：零向量退化 / code 03, degenerate zero vector
    RETURN;
END_IF

// 段 5｜圆均值求解：ATAN2 于 (fxSum, fySum)，fR ≥ 1E-6 保证不会落在 (0,0) 点
//      segment 5, the mean via atan2, the magnitude gate keeps the point off the origin
fMean := ATAN2(fySum, fxSum) / CMC_DEG2RAD;             // 弧度回角度 [°] / radians back to degrees [deg]

// 段 6｜归一 [0,360)：条件加减搬区间，禁负取模 / segment 6, normalise to [0,360) by conditional add or subtract
IF fMean < 0.0 THEN
    fMean := fMean + CMC_DEG_TURN;                      // 负半区搬上去（ATAN2 值域 ±180，一次即够）/ move the negative half up
END_IF
IF fMean >= CMC_DEG_TURN THEN
    fMean := fMean - CMC_DEG_TURN;                      // 满圈搬下来（数值抖动防线）/ bring a full turn down
END_IF

// 段 7｜出口 / segment 7, exit
FC_DL_CircularMeanCalc := fMean;                        // 发布圆均值 [°] / publish the circular mean [deg]
bValid := TRUE;                                         // 结果可用 / the result is usable
END_FUNCTION

(* ---- FC_DL_ConductivityTempComp.st ---- *)
(*
  ==================================================================
  组件名 Component  : FC_DL_ConductivityTempComp
  分类   Category   : DL_MathData
  复杂度 Complexity  : 中
  版本   Version    : 1.0.0
  功能   Purpose    : 电导率温度补偿（参考温归一）。κ_ref = κ_T / (1 +
                      α(T − T_ref))，α 为温度系数 [%每摄氏度]，域 [0,5]；
                      测温域 [0,60] 摄氏度，越域钳位并置 bOutOfRange（信息级
                      超域标志）；补偿分母下限闸防除零与负分母。OSCAT
                      Building 水质域公开语义 clean-room。
  来源   Source     : T1-2-oscat-building（水质域公开语义）
  溯源   Origin     : 线性温度补偿公式为公开水质工程语义，clean-room 自研
                      实现，未复制 OSCAT 或任何厂商私有库源码。
  平台   Platform   : 纯 IEC 61131-3，CODESYS / TwinCAT / InoProShop 通用
  分工声明 Split     : 与 FC_DL_PhCompensation 分工——后者做 pH 温度补偿，
                      本件做电导率参考温归一。
  作者   Author     : 道莅代码库 · PLC 编程专家（R59）
  ------------------------------------------------------------------
  边界 Boundary     :
                      一 非有限入参闸（自反双判据，三参数全覆盖）：命中置
                         bError，输出安全侧零（四段式 R45）；
                      二 测温域 [0,60] 与系数域 [0,5] 越域钳位并置
                         bOutOfRange / bClamped（信息级，单点回夹）；
                      三 除零与负分母闸：分母 < 0.1 置 bError（防 1+αΔT
                         趋零或变负，含负绝对温差场景）；
                      四 无全局变量、无外部变量声明、无物理地址寻址。
  修订记录 Revision  :
    2026-11-21  v1.0.0  R59 首版（批 4 · 序号 17）
  ==================================================================
*)

FUNCTION FC_DL_ConductivityTempComp : BOOL
VAR_INPUT
    fCondRaw  : LREAL := 0.0; // 电导率实测值 [微西门子每厘米] / the measured conductivity [microsiemens per centimeter]
    fTempC    : LREAL := 25.0; // 水样温度 [摄氏度]，域 [0,60] / the sample temperature [degree celsius]
    fAlphaPct : LREAL := 2.0;  // 温度系数 [%每摄氏度]，域 [0,5] / the temperature coefficient [percent per degree celsius]
    fRefTempC : LREAL := 25.0; // 参考温度 [摄氏度] / the reference temperature [degree celsius]
END_VAR
VAR_OUTPUT
    fCondRef    : LREAL := 0.0; // 参考温归一电导率 [微西门子每厘米] / the normalized conductivity [microsiemens per centimeter]
    bValid      : BOOL := FALSE; // 结果可用标志 [-] / the result usable flag
    bOutOfRange : BOOL := FALSE; // 测温越域标志（信息级）[-] / the temperature out of range flag, informational
    bClamped    : BOOL := FALSE; // 系数越域钳位（信息级）[-] / the coefficient clamp, informational
    bError      : BOOL := FALSE; // 故障标志（非有限或分母退化）[-] / the fault flag
END_VAR
VAR CONSTANT
    DL_CTC_TMIN  : LREAL := 0.0;  // 测温域下界 [摄氏度] / the temperature floor
    DL_CTC_TMAX  : LREAL := 60.0; // 测温域上界 [摄氏度] / the temperature ceiling
    DL_CTC_AMIN  : LREAL := 0.0;  // 系数域下界 [%每摄氏度] / the coefficient floor
    DL_CTC_AMAX  : LREAL := 5.0;  // 系数域上界 [%每摄氏度] / the coefficient ceiling
    DL_CTC_DENMIN: LREAL := 0.1;  // 补偿分母下限 [无量纲] / the denominator floor
END_VAR
VAR
    lrT    : LREAL; // 测温工作量（钳后）[摄氏度] / the clamped temperature work value
    lrAlp  : LREAL; // 系数工作量（钳后）[%每摄氏度] / the clamped coefficient work value
    lrDen  : LREAL; // 补偿分母工作量 [无量纲] / the denominator work value
    bFin   : BOOL;  // 入参有限工作量 [-] / the input finiteness work flag
END_VAR

// 段 1｜返回值与输出预置（四段式第一段，R45）/ segment 1, preset the return and the outputs
FC_DL_ConductivityTempComp := FALSE; // 受理预置假 / preset the accepted false
fCondRef := 0.0; // 输出预置零 / preset the output zero
bValid := FALSE; // 有效预置假 / preset the valid false
bOutOfRange := FALSE; // 越域预置假 / preset the range flag false
bClamped := FALSE; // 钳位预置假 / preset the clamp false
bError := FALSE; // 故障预置假 / preset the fault false

// 段 2｜非有限入参闸（三参数自反双判据全覆盖，R79）/ segment 2, the non finite gate
bFin := (fCondRaw = fCondRaw) AND ((fCondRaw - fCondRaw) = (fCondRaw - fCondRaw)) // 电导率有限 / the conductivity finite
    AND (fTempC = fTempC) AND ((fTempC - fTempC) = (fTempC - fTempC)) // 测温有限 / the temperature finite
    AND (fAlphaPct = fAlphaPct) AND ((fAlphaPct - fAlphaPct) = (fAlphaPct - fAlphaPct)) // 系数有限 / the coefficient finite
    AND (fRefTempC = fRefTempC) AND ((fRefTempC - fRefTempC) = (fRefTempC - fRefTempC)); // 参考温有限 / the reference finite
IF NOT bFin THEN // 非有限命中 / a non finite hit
    bError := TRUE; // 置故障（纪律②）/ raise the fault
    RETURN; // 早退 / return early
END_IF

// 段 3｜域钳制（测温越域置 bOutOfRange，系数钳位置 bClamped，边界二）/ segment 3, the domain clamps
lrT := fTempC; // 装测温 / load the temperature
IF (lrT < DL_CTC_TMIN) OR (lrT > DL_CTC_TMAX) THEN // 测温越域 / the temperature out of range
    bOutOfRange := TRUE; // 置超域标志（信息级）/ raise the out of range flag
    IF lrT < DL_CTC_TMIN THEN // 下越界 / below the floor
        lrT := DL_CTC_TMIN; // 钳到下界 / clamp to the floor
    ELSE // 上越界 / above the ceiling
        lrT := DL_CTC_TMAX; // 钳到上界 / clamp to the ceiling
    END_IF
END_IF
lrAlp := fAlphaPct; // 装系数 / load the coefficient
IF lrAlp < DL_CTC_AMIN THEN // 系数下钳 / clamp the coefficient down
    lrAlp := DL_CTC_AMIN; // 夹到零 / clamp to the floor
    bClamped := TRUE; // 信息级 / informational
ELSIF lrAlp > DL_CTC_AMAX THEN // 系数上钳 / clamp the coefficient up
    lrAlp := DL_CTC_AMAX; // 夹到上限 / clamp to the ceiling
    bClamped := TRUE; // 信息级 / informational
END_IF

// 段 4｜补偿计算（分母下限闸防除零与负分母，边界三）/ segment 4, the compensation with the denominator gate
lrDen := 1.0 + ((lrAlp / 100.0) * (lrT - fRefTempC)); // 补偿分母 / the denominator
IF lrDen < DL_CTC_DENMIN THEN // 分母退化闸（除零与负分母双防）/ the degenerate denominator gate
    bError := TRUE; // 置故障（纪律②）/ raise the fault
    RETURN; // 早退 / return early
END_IF
fCondRef := fCondRaw / lrDen; // 参考温归一（除子已闸）/ the normalization, divided by the gated denominator
bValid := TRUE; // 结果可用 / the result usable
FC_DL_ConductivityTempComp := TRUE; // 受理 / accept
END_FUNCTION

(* ---- FC_DL_CosDeg.st ---- *)
(*==============================================================================
 * 名称 : FC_DL_CosDeg —— 角度制余弦（度入参，弧度内部换算）
 * 分类 / 前缀 / 版本 : DL_MathData / FC_DL_ / 1.0.0
 * 溯源 : 开源语义参考（OSCAT/AixOCAT 族，MIT）或 clean-room IEC 实现，未复制源码
 * 平台 : 纯 IEC 61131-3
 * 功能说明 : 返回 cos(fDeg)：内部换算弧度 fDeg * PI / 180 后调用标准 COS，
 *            PI 取 LREAL 字面量 3.14159265358979323846（双精度最近舍入）。
 *            边界处理：输入非有限（NaN：f<>f；±Inf：(f-f)<>(f-f)）置 eErr
 *            返回 0.0；|fDeg|>1.0E12 时大角换算精度塌陷，同置 eErr 返回 0.0。
 * 错误码 : 16#0001_1B0A = 输入非有限（NaN/±Inf）或角度量超安全量程 ±1.0E12
 *          eErr=0 且 bValid=TRUE 表示返回值可用
 * 状态机 : R6 标注 N/A（纯函数无顺序状态，以本节替代 ELSE 兜底）
 * 红线 : R1/R2/R3 ✓ 零全局/零IO/纯IEC ｜ R4 ✓ 非有限拦截/量程防护 ｜ R10 ✓ 标准转换 ｜ R11 ✓ 分号收尾 ｜ R15 ✓ 无保留字撞名
 * 修订记录 : 2026-11-23 v1.0.0 首次入库（R76）
 *============================================================================*)
FUNCTION FC_DL_CosDeg : LREAL
VAR_INPUT
    fDeg : LREAL;    // 输入角 [度] / input angle in degrees
END_VAR
VAR_OUTPUT
    eErr   : UDINT;    // 故障码，0=正常，1B0A=输入非有限或超量程 / error code
    bError : BOOL;     // TRUE=本件发生故障 / TRUE when fault occurred
    bValid : BOOL;     // TRUE=返回值可用 / TRUE when return value is usable
END_VAR

FC_DL_CosDeg := 0.0;                         // 返回值预设 0.0 / preset return to zero
eErr   := 16#0000_0000;                      // 故障码清零 / clear error code
bError := FALSE;                             // 故障标志清零 / clear error flag
bValid := TRUE;                              // 预设输出可用 / preset valid flag

IF (fDeg <> fDeg) OR ((fDeg - fDeg) <> (fDeg - fDeg))    // NaN 或 ±Inf / NaN or infinite
   OR (ABS(fDeg) > 1.0E12) THEN              // 超安全量程（精度塌陷防护）/ beyond safe range
    eErr   := 16#0001_1B0A;                  // 置故障码 / set error code
    bError := TRUE;                          // 置故障标志 / set error flag
    bValid := FALSE;                         // 返回值不可用 / return not usable
    RETURN;                                  // 返回 0.0 / return zero
END_IF

FC_DL_CosDeg := COS(fDeg * 3.14159265358979323846 / 180.0);    // 度转弧度后取余弦 / degrees to radians, then cosine

END_FUNCTION

(* ---- FC_DL_CosEx.st ---- *)
(*
    FC_DL_CosEx —— 余弦防御包装（与 SinEx 同一 2π 归约策略 + 非有限拦截 + 超大角度降级）
    ------------------------------------------------------------------
    分类      : DL_MathData / Math-Trig
    前缀      : FC_DL_
    版本      : 1.0.0
    溯源      : IEC 61131-3 标准语义的道莅防御性实现
                （内部委托平台内建函数，外围统一错误码/钳位/双语文档；
                  未复制任何闭源厂商源码，参考实现仅限 MIT/Apache 许可）
    平台      : 纯 IEC 61131-3，CODESYS / TwinCAT / InoProShop 通用
    作者      : 道莅代码库 · PLC编程专家（R15）
    ------------------------------------------------------------------
    功能说明  : 求输入弧度的余弦值，归约策略与 FC_DL_SinEx 完全一致。
                入口先做非有限拦截（NaN/Inf 返回 0.0 并置 16#0001_0168）；随后按
                2π 做周期归约，商取 FLOOR 语义，商绝对值 < 2.0E9 保证
                DINT 转换不溢出；超大角度（绝对值 > 1.0E12 或商超 DINT
                安全域）置 16#0001_0168、bValid=FALSE 降级但仍继续计算；域内委托
                内建 COS，结果再做 NaN 复检兜底，全程不输出 NaN/Inf。
    错误码    : 0000 正常 / 16#0001_0168 入参越界（非有限输入或超大角度降级，已归零/降级可用）
    修订记录  : 2026-11-16 v1.0.0 首次入库（R15）
*)
FUNCTION FC_DL_CosEx : LREAL
VAR_INPUT
    lrRad : LREAL; // 输入角度 [rad]，任意有限弧度值 / input angle [rad], any finite radian value
END_VAR
VAR_OUTPUT
    eErr : UDINT; // 错误码，0=正常，1=入参越界（非有限或超大角度） / error id, 0=ok, 1=input out of domain (non-finite or super-large angle)
    bError   : BOOL; // 是否出错，eErr 非 0 时为 TRUE / error flag, TRUE when eErr is nonzero
    bValid   : BOOL; // 输出是否有效可用，超大角度降级时为 FALSE / output valid, FALSE for degraded super-large angle
END_VAR
VAR
    lrQ   : LREAL; // 周期商 [周期数]，输入角除以 2π / cycle quotient [cycles], input divided by two pi
    nCyc  : DINT; // 归约周期数 [周期数]，FLOOR 语义整数 / reduction cycle count [cycles], integer with floor semantics
    lrRed : LREAL; // 归约后弧度 [rad]，域约至 0 到 2π / reduced angle [rad], bounded to 0 to 2 pi
END_VAR
VAR CONSTANT
    DL_CS_MAXREAL : LREAL := 1.7976931348623157E308; // 双精度有限极值 [rad]，超界判无穷 / double precision finite max [rad], beyond treated as infinity
    DL_CS_TWOPI   : LREAL := 6.283185307179586; // 圆周率两倍 [rad]，归约模数 / two pi [rad], reduction modulus
    DL_CS_BIG     : LREAL := 1.0E12; // 超大角度阈值 [rad]，超过判降级 / super-large angle threshold [rad], beyond degraded
    DL_CS_QMAX    : LREAL := 2.0E9; // 周期商安全域 [周期数]，保证 DINT 转换不溢出 / quotient safe bound [cycles], keeps DINT conversion overflow-free
    DL_CS_EPS     : LREAL := 1.0E-9; // 浮点容差 [无量纲] / floating point tolerance [dimensionless]
END_VAR

// 段 1｜返回值与错误状态预置，任何早退路径不留脏码 / segment 1, preset return value and error states
FC_DL_CosEx := 0.0; // 返回值预置安全值 0.0 / preset return to safe value 0.0
eErr    := 16#0000_0000; // 错误码预置正常 / preset error id to ok
bError      := FALSE; // 错误标志预置无错 / preset error flag to FALSE
bValid      := TRUE; // 有效标志预置可用 / preset valid flag to TRUE

// 段 2｜非有限拦截：NaN 用自不等判据，无穷用超极值判据 / segment 2, non-finite interception
IF (lrRad <> lrRad) OR (lrRad > DL_CS_MAXREAL) OR (lrRad < -DL_CS_MAXREAL) THEN
    eErr := 16#0001_0168; // 信息级：输入非有限，已归零 / informational, non-finite input, zeroed
    bError   := TRUE; // 置错误标志 / raise error flag
    bValid   := FALSE; // 输出不可用 / output invalid
    RETURN; // 返回预置安全值 0.0 / return preset safe value 0.0
END_IF

// 段 3｜2π 周期归约（FLOOR 语义）：商超 DINT 安全域则跳过归约原值直通 / segment 3, two-pi reduction with floor semantics, skipped when quotient exceeds the DINT safe bound
lrQ := lrRad / DL_CS_TWOPI; // 周期商 [周期数] / cycle quotient [cycles]
IF ABS(lrQ) < DL_CS_QMAX THEN
    nCyc := TRUNC(lrQ); // 向零截取周期数 / truncate quotient toward zero
    IF (lrQ < 0.0) AND (ABS(lrQ - DINT_TO_LREAL(nCyc)) > DL_CS_EPS) THEN
        nCyc := nCyc - 1; // 负非整数商补一，落实 FLOOR 语义 / decrement for negative non-integer quotient to enforce floor semantics
    END_IF
    lrRed := lrRad - DL_CS_TWOPI * DINT_TO_LREAL(nCyc); // 归约后弧度 [rad] / reduced angle [rad]
ELSE
    lrRed := lrRad; // 商超安全域，放弃归约原值直通 / quotient beyond safe bound, reduction skipped
END_IF

// 段 4｜超大角度精度闸：置 16#0001_0168 降级但继续计算 / segment 4, super-large angle precision gate, degraded with code 1 but computation continues
IF (ABS(lrRad) > DL_CS_BIG) OR (ABS(lrQ) >= DL_CS_QMAX) THEN
    eErr := 16#0001_0168; // 信息级：超大角度，精度不可保证 / informational, super-large angle, precision not guaranteed
    bError   := TRUE; // 置错误标志 / raise error flag
    bValid   := FALSE; // 降级输出，需上层注意 / degraded output, upper layer attention required
END_IF

// 段 5｜委托内建 COS + 结果 NaN 复检兜底 / segment 5, delegation to built-in COS with result NaN recheck
FC_DL_CosEx := COS(lrRed); // 委托内建 COS 内核，不自实现三角内核 / delegate to built-in COS kernel
IF FC_DL_CosEx <> FC_DL_CosEx THEN
    FC_DL_CosEx := 0.0; // 兜底安全值 / bottom-line safe value
    IF eErr = 16#0000_0000 THEN
        eErr := 16#0001_0168; // 首事件优先置码 / first-event priority code
        bError   := TRUE; // 置错误标志 / raise error flag
        bValid   := FALSE; // 输出不可用 / output invalid
    END_IF
END_IF
END_FUNCTION

(* ---- FC_DL_CpkCalc.st ---- *)
// =====================================================================
// FC_DL_CpkCalc.st
// 过程能力指数计算纯函数 (Cp/Cpu/Cpl/Cpk) SPC 自研 T2-8
// Process capability index calculation pure function
// 码位: 16#0001_0480 ~ 16#0001_0484 (本件独占 5 槽)
// 修改记录: R29 初版 (按 DISPATCH_R29 序 2)
// =====================================================================
FUNCTION FC_DL_CpkCalc : BOOL
VAR_INPUT
    bEnable      : BOOL   := TRUE;      // 使能 / Enable
    fMean        : REAL   := 0.0;       // 样本均值（工程单位）/ Sample mean [unit]
    fSigma       : REAL   := 0.0;       // 样本标准差 ≥0（同单位）/ Sample sigma [unit]
    fUsl         : REAL   := 100.0;     // 规格上限 / Upper spec limit [unit]
    fLsl         : REAL   := 0.0;       // 规格下限 / Lower spec limit [unit]
    uSampleCount : UDINT  := 0;         // 样本数 / Sample count
    uSampleMin   : UDINT  := 25;        // 最小样本数 5~1000 / Minimum sample count
    fSigmaMin    : REAL   := 1.0E-6;    // σ 下限 >0（退化判据）/ Sigma floor [unit]
    fCpkMin      : REAL   := 1.33;      // 合格门限 0.5~3.0 / Capability threshold [-]
END_VAR
VAR_OUTPUT
    fCp          : REAL;                // 潜在能力 / Potential capability [-]
    fCpu         : REAL;                // 上侧能力 / Upper capability [-]
    fCpl         : REAL;                // 下侧能力 / Lower capability [-]
    fCpk         : REAL;                // 实际能力 / Actual capability [-]
    bValid       : BOOL;                // 结论有效 / Result valid
    bCapable     : BOOL;                // 达门限 / Capable
    eErr         : UDINT;               // 错误码 / Error code
END_VAR
VAR
    fSigmaClamp  : REAL;                // 钳下限后的 σ / Clamped sigma [unit]
    fThreeSig    : REAL;                // 3σ 分母 / 3-sigma denominator [unit]
    fSixSig      : REAL;                // 6σ 分母 / 6-sigma denominator [unit]
    fCpkMinSafe  : REAL;                // 非有限兜底后的门限 / Sanitized threshold [-]
END_VAR

// ---------------------------------------------------------------------
// 代码位表（本件独占，勿复用）:
//   16#0001_0480 信息 计算完成且结论有效
//   16#0001_0481 故障 fMean/fSigma/fUsl/fLsl 非有限，或 fSigma < 0
//   16#0001_0482 故障 fUsl ≤ fLsl（组态错），或 fSigmaMin ≤ 0
//   16#0001_0483 信息 退化：fSigma < fSigmaMin → Cp/Cpk 置 999.0 哨兵、bValid=FALSE
//   16#0001_0484 信息 样本不足：uSampleCount < uSampleMin → 输出全 0、bValid=FALSE
// ---------------------------------------------------------------------

// 默认输出清零 / Default outputs cleared
fCp      := 0.0;      // Cp 清零 / Reset Cp
fCpu     := 0.0;      // Cpu 清零 / Reset Cpu
fCpl     := 0.0;      // Cpl 清零 / Reset Cpl
fCpk     := 0.0;      // Cpk 清零 / Reset Cpk
bValid   := FALSE;    // 结论无效 / Invalid by default
bCapable := FALSE;    // 未达门限 / Not capable by default
eErr     := 16#0001_0480;  // 预置正常码 / Preset normal code

IF NOT bEnable THEN
    // 使能关闭：输出保持 0，不置故障 / Disabled: outputs zero, no fault
    RETURN;   // 直接返回 / Return
END_IF

// ---- 非有限闸 / Finite guard ----
IF (fMean <> fMean) OR (ABS(fMean) >= 1.0E12)
   OR (fSigma <> fSigma) OR (ABS(fSigma) >= 1.0E12)
   OR (fUsl <> fUsl) OR (ABS(fUsl) >= 1.0E12)
   OR (fLsl <> fLsl) OR (ABS(fLsl) >= 1.0E12) THEN
    eErr := 16#0001_0481;  // 故障：输入非有限 / Fault: non-finite input
    RETURN;                // 输出保持 0 / Outputs stay zero
END_IF

// ---- σ 负值判 / Negative sigma fault ----
IF fSigma < 0.0 THEN
    eErr := 16#0001_0481;  // 故障：σ < 0 / Fault: sigma negative
    RETURN;                // 输出保持 0 / Outputs stay zero
END_IF

// ---- 组态错闸 / Configuration fault ----
IF (fUsl <= fLsl) OR (fSigmaMin <= 0.0) THEN
    eErr := 16#0001_0482;  // 故障：规格区间或 σ 下限非法 / Fault: invalid spec or sigma floor
    RETURN;                // 输出保持 0 / Outputs stay zero
END_IF

// ---- 门限脏值兜底（不置错）/ Sanitize dirty threshold without fault ----
fCpkMinSafe := fCpkMin;                     // 先原样采用 / Adopt as-is first
IF (fCpkMin <> fCpkMin) OR (ABS(fCpkMin) >= 1.0E12) THEN
    fCpkMinSafe := 1.33;                    // 兜底 1.33 / Fallback 1.33
END_IF

// ---- 样本数不足 → 输出全 0 不给结论 / Insufficient samples ----
IF uSampleCount < uSampleMin THEN
    eErr := 16#0001_0484;  // 信息级：样本不足 / Info: insufficient samples
    RETURN;                // 输出保持 0，bValid=FALSE / Outputs zero, invalid
END_IF

// ---- 退化判：σ < σMin → 哨兵 999.0，不得报除零 / Degenerate sigma sentinel ----
IF fSigma < fSigmaMin THEN
    fCp    := 999.0;        // Cp 哨兵 / Cp sentinel
    fCpk   := 999.0;        // Cpk 哨兵 / Cpk sentinel
    bValid := FALSE;        // 结论无效 / Invalid
    eErr   := 16#0001_0483; // 信息级：退化 / Info: degenerate
    RETURN;                 // 直接返回 / Return
END_IF

// ---- 先钳 σ 下限再除，杜绝 3σ/6σ 除零热点 / Clamp sigma before division ----
IF fSigma < fSigmaMin THEN
    fSigmaClamp := fSigmaMin;   // 保险钳位（理论上不可达）/ Defensive clamp
ELSE
    fSigmaClamp := fSigma;      // 正常 σ / Normal sigma
END_IF
fThreeSig := 3.0 * fSigmaClamp; // 3σ 分母 / 3-sigma denominator
fSixSig   := 6.0 * fSigmaClamp; // 6σ 分母 / 6-sigma denominator

// ---- 四项能力指数 / Four capability indices ----
fCp  := (fUsl - fLsl) / fSixSig;   // Cp = (USL-LSL)/(6σ) / Potential capability
fCpu := (fUsl - fMean) / fThreeSig; // Cpu = (USL-μ)/(3σ) / Upper capability
fCpl := (fMean - fLsl) / fThreeSig; // Cpl = (μ-LSL)/(3σ) / Lower capability

// Cpk = MIN(Cpu, Cpl)，负值照实输出禁止钳零 / Cpk as-is, no clamping
IF fCpu <= fCpl THEN
    fCpk := fCpu;   // 取上侧较小值 / Take upper
ELSE
    fCpk := fCpl;   // 取下侧较小值 / Take lower
END_IF

// ---- 结论与达标判 / Validity and capability verdict ----
bValid   := TRUE;              // 结论有效 / Valid
bCapable := (fCpk >= fCpkMinSafe);  // 达门限判 / Threshold verdict

// 正常完成，返回 TRUE / Normal completion
FC_DL_CpkCalc := TRUE;         // 函数返回值 / Function result

END_FUNCTION

(* ---- FC_DL_CpkIndex.st ---- *)
(*
    FC_DL_CpkIndex —— 过程能力指数 Cp / Cpk
    ------------------------------------------------------------------
    分类      : DL_MathData / Statistics
    前缀      : FC_DL_
    版本      : 1.0.0
    溯源      : 自研（Cp / Cpk 为公开统计定义）；ISO 22400-2 质量口径仅作术语参考
                （T2-8 次源，不复制任何条款文本）；
                clean-room 重写，未复制任何闭源厂商源码，参考实现仅限 MIT/Apache 许可
    平台      : 纯 IEC 61131-3，CODESYS V3.5+ / TwinCAT 3 / InoProShop 通用
    作者      : 道莅代码库 · PLC编程专家（R18）
    ------------------------------------------------------------------
    功能说明  : 由样本数组算 Cp、Cpk、均值与样本标准差（n-1 分母），供质量工站实时判
                工序能力（Cpk 小于 1.33 报警）；与 SignalStatistics 的分界是本件以规格
                限为输入、以能力指数为出口，不做通用统计量集合；
                防御链：规格限合法性闸 → 样本数闸 → 非有限样本逐点剔除 → σ 近零饱和闸
                → 六倍σ除号闸，每一闸都在除法之前；
                累加与方差用 LREAL 中间量，64 点大值平方不会溢出（R10 同纪律）。
    错误码    : 16#0001_0243 σ 近零，Cp / Cpk 已按饱和上限输出（常数样本，合法工况）——信息级，不置故障
                16#0001_0244 预留禁用（信息级，不得挪用）
                16#0001_031B 有效样本数不足（小于 2），无法计算——故障级，返回 0
                16#0001_031C 规格限非法（上限不大于下限）——故障级，返回 0
                16#0001_031D 预留禁用（故障级，不得挪用）
    码位总账  : 16#0001_0243 用 / 16#0001_0244 预留 ｜ 16#0001_031B 用 / 16#0001_031C 用 / 16#0001_031D 预留
    状态机    : N/A —— 纯函数无顺序状态机，无 CASE 可写，非法状态不可能出现
    采样约定  : 纯组合函数，无定时器、无内部驻留状态；样本窗由调用方滚动填充，
                本件按 uCount 指定的前缀区间读取，绝不读取未填充的尾部。
    修订记录  : 2026-11-16 v1.0.0 首次入库（R18）
*)
FUNCTION FC_DL_CpkIndex : REAL
VAR_INPUT
    afSample : ARRAY[0..63] OF REAL;           // 样本数组，有效项 0~uCount-1 [用户单位] / sample array, valid items 0~uCount-1 [user unit]
    uCount   : UINT := 0;                      // 样本数 [个]，范围 2~64 / sample count [item], range 2~64
    fLsl     : REAL := 0.0;                    // 规格下限 [用户单位] / lower specification limit [user unit]
    fUsl     : REAL := 1.0;                    // 规格上限，必须大于下限 [用户单位] / upper specification limit, must exceed the lower one [user unit]
    fCpkSat  : REAL := 10.0;                   // Cpk 饱和上限（σ 近零时输出此值）[无量纲]，范围 1.0~100.0 / Cpk saturation cap [dimensionless], range 1.0~100.0
END_VAR
VAR_OUTPUT
    fCp        : REAL;                         // 潜在能力指数（不含偏移）[无量纲] / potential capability index without offset [dimensionless]
    fCpk       : REAL;                         // 实际能力指数，返回值的镜像 [无量纲] / actual capability index, mirror of the return value [dimensionless]
    fMean      : REAL;                         // 样本均值 [用户单位] / sample mean [user unit]
    fSigma     : REAL;                         // 样本标准差（n-1 分母）[用户单位] / sample standard deviation with n-1 denominator [user unit]
    eErr       : UDINT;                        // 错误码，0=正常 / error id, 0=ok
    bError     : BOOL;                         // 故障标志，eErr 为故障级时 TRUE / error flag, TRUE on fault-level eErr
    bValid     : BOOL;                         // 结果是否可用 / result usable flag
    bSaturated : BOOL;                         // 因 σ 近零而饱和 / saturated because sigma is near zero
END_VAR
VAR
    uIdx     : UINT;                           // 样本游标 [个] / sample cursor [item]
    uValidN  : UINT;                           // 剔除后有效样本数 [个] / valid sample count after removal [item]
    uKicked  : UINT;                           // 被剔除的非有限样本数 [个] / non-finite samples removed [item]
    fSum     : LREAL;                          // 样本和，LREAL 中间量防溢出 [用户单位] / sample sum, LREAL intermediate against overflow [user unit]
    fSumSq   : LREAL;                          // 偏差平方和，LREAL 中间量防溢出 [用户单位平方] / sum of squared deviations, LREAL intermediate [user unit squared]
    fDev     : REAL;                           // 单个样本偏差 [用户单位] / single sample deviation [user unit]
    fMeanL   : LREAL;                          // 均值 LREAL 中间量 [用户单位] / mean as LREAL intermediate [user unit]
    fVar     : LREAL;                          // 样本方差（n-1 分母）[用户单位平方] / sample variance with n-1 denominator [user unit squared]
    fSpan    : REAL;                           // 六倍标准差，Cp 分母 [用户单位] / six sigma span, the Cp denominator [user unit]
    fUpper   : REAL;                           // 上侧能力 [无量纲] / upper side capability [dimensionless]
    fLower   : REAL;                           // 下侧能力 [无量纲] / lower side capability [dimensionless]
    bNonFin  : BOOL;                           // 单个样本非有限判定标志 / single sample non-finite flag
END_VAR
VAR CONSTANT
    DL_CPK_MAX_N     : UINT := 64;             // 样本数上限 [个] / sample count upper bound [item]
    DL_CPK_MIN_N     : UINT := 2;              // 样本数下限，n 小于 2 时 σ 无定义 [个] / sample count lower bound, sigma is undefined below two [item]
    DL_CPK_LAST_IDX  : UINT := 63;             // 样本数组末索引 [个] / last sample index [item]
    DL_FLOAT_EPS     : REAL := 1.0E-6;         // 浮点判等容差 [用户单位] / float equality tolerance [user unit]
    DL_CPK_INF_GUARD : REAL := 4.0E38;         // 非有限幅值判定阈值 [用户单位] / non-finite magnitude guard [user unit]
    DL_CPK_SIGMA_K    : REAL := 3.0;           // 单侧三倍标准差 [无量纲] / three sigma per side [dimensionless]
    DL_CPK_SIGMA_6    : REAL := 6.0;           // 双侧六倍标准差 [无量纲] / six sigma over both sides [dimensionless]
    DL_CPK_SAT_MIN    : REAL := 1.0;           // 饱和上限下限 [无量纲] / lower bound of the saturation cap [dimensionless]
    DL_CPK_SAT_MAX    : REAL := 100.0;         // 饱和上限上限 [无量纲] / upper bound of the saturation cap [dimensionless]
    DL_CPK_ZERO       : REAL := 0.0;           // 零值常量，避免裸字面量 [无量纲] / zero constant, avoids a bare literal [dimensionless]
    DL_CPK_N1         : UINT := 1;             // n-1 分母的减数 [个] / subtrahend of the n-1 denominator [item]
END_VAR

// 段 1｜返回值与输出预置 / segment 1, preset return value and outputs
FC_DL_CpkIndex := DL_CPK_ZERO;                 // 故障缺省返回 0 / fault default returns zero
fCp := DL_CPK_ZERO;                            // Cp 预置 0 / preset Cp to zero
fCpk := DL_CPK_ZERO;                           // Cpk 预置 0 / preset Cpk to zero
fMean := DL_CPK_ZERO;                          // 均值预置 0 / preset the mean to zero
fSigma := DL_CPK_ZERO;                         // 标准差预置 0 / preset sigma to zero
eErr := 0;                                     // 预置无错误 / preset no error
bError := FALSE;                               // 预置无故障 / preset no fault
bValid := FALSE;                               // 预置结果不可用 / preset unusable
bSaturated := FALSE;                           // 预置未饱和 / preset not saturated
uValidN := 0;                                  // 有效样本数清零 / clear the valid count
uKicked := 0;                                  // 剔除数清零 / clear the removed count
fSum := 0.0;                                   // 求和清零 / clear the sum
fSumSq := 0.0;                                 // 平方和清零 / clear the squared sum

// 段 2｜饱和上限闸：越域即钳位，符号方向写进注释 / segment 2, saturation cap gate
IF (fCpkSat < DL_CPK_SAT_MIN) OR (fCpkSat > DL_CPK_SAT_MAX) THEN
    fCpkSat := MIN(MAX(fCpkSat, DL_CPK_SAT_MIN), DL_CPK_SAT_MAX); // 双侧钳位到 1.0~100.0 / clamp both sides into 1.0~100.0
END_IF

// 段 3｜规格限闸：上限不大于下限即非法，容差内视为相等同样非法 / segment 3, specification limit gate
IF (fUsl - fLsl) <= DL_FLOAT_EPS THEN
    eErr := 16#0001_031C;                      // 规格限非法故障码 / illegal specification limit fault id
    bError := TRUE;                            // 置故障标志 / raise the error flag
    RETURN;                                    // 故障级提前返回 / early return on fault
END_IF

// 段 4｜样本数闸：先判界再索引 / segment 4, sample count gate before any indexing
IF (uCount < DL_CPK_MIN_N) OR (uCount > DL_CPK_MAX_N) THEN
    eErr := 16#0001_031B;                      // 样本数不足或越界故障码 / insufficient or out of range sample count fault id
    bError := TRUE;                            // 置故障标志 / raise the error flag
    RETURN;                                    // 故障级提前返回 / early return on fault
END_IF

// 段 5｜第一遍：剔除非有限样本并求和 / segment 5, first pass removes non-finite samples and sums the rest
FOR uIdx := 0 TO uCount - 1 DO
    bNonFin := (afSample[uIdx] <> afSample[uIdx])
            OR (afSample[uIdx] > DL_CPK_INF_GUARD)
            OR (afSample[uIdx] < -DL_CPK_INF_GUARD); // 非有限判定 / non-finite check
    IF bNonFin THEN
        uKicked := uKicked + 1;                // 剔除计数，NaN 参与求和会污染全部结果 / count the removal, a NaN would poison the whole sum
    ELSE
        fSum := fSum + afSample[uIdx];         // LREAL 累加 / accumulate in LREAL
        uValidN := uValidN + 1;                // 有效样本计数 / count the valid sample
    END_IF
END_FOR
IF uValidN < DL_CPK_MIN_N THEN
    eErr := 16#0001_031B;                      // 剔除后仍不足两个有效样本 / still fewer than two valid samples after removal
    bError := TRUE;                            // 置故障标志 / raise the error flag
    RETURN;                                    // 故障级提前返回 / early return on fault
END_IF

// 段 6｜均值与第二遍方差（两遍法比一次式 sumsq 数值稳定）/ segment 6, mean and second pass variance
fMeanL := fSum / UINT_TO_LREAL(uValidN);       // 分母由段 4 与段 5 保证不小于 2，显式升位转换 / the denominator is at least two thanks to the gates above, widened explicitly
fMean := LREAL_TO_REAL(fMeanL);                // 均值对外输出 / publish the mean
FOR uIdx := 0 TO uCount - 1 DO
    bNonFin := (afSample[uIdx] <> afSample[uIdx])
            OR (afSample[uIdx] > DL_CPK_INF_GUARD)
            OR (afSample[uIdx] < -DL_CPK_INF_GUARD); // 剔除样本不参与方差 / removed samples never enter the variance
    IF NOT bNonFin THEN
        fDev := afSample[uIdx] - fMean;        // 偏差 / deviation from the mean
        fSumSq := fSumSq + REAL_TO_LREAL(fDev) * REAL_TO_LREAL(fDev); // LREAL 乘方防溢出 / square in LREAL against overflow
    END_IF
END_FOR
fVar := fSumSq / UINT_TO_LREAL(uValidN - DL_CPK_N1); // n-1 分母，无偏估计，显式升位 / unbiased estimate with the n-1 denominator, widened explicitly
IF fVar < 0.0 THEN
    fVar := 0.0;                               // 数值噪声可能产生极小负值，钳到 0 再开方 / numerical noise may go slightly negative, clamp before the root
END_IF
fSigma := LREAL_TO_REAL(SQRT(fVar));           // 样本标准差 / sample standard deviation

// 段 7｜σ 近零饱和闸：常数样本是合法工况，只置信息码不置故障 / segment 7, sigma near zero saturation gate
IF fSigma <= DL_FLOAT_EPS THEN
    fCp := fCpkSat;                            // 潜在能力按饱和上限输出 / potential capability saturates
    fCpk := fCpkSat;                           // 实际能力按饱和上限输出 / actual capability saturates
    FC_DL_CpkIndex := fCpkSat;                 // 返回值同为饱和上限 / the return value follows the cap
    bSaturated := TRUE;                        // 标记饱和 / flag the saturation
    bValid := TRUE;                            // 饱和值是可用结果 / the saturated value is usable
    eErr := 16#0001_0243;                      // 饱和提示（信息级不置故障）/ saturation hint, info level never raises a fault
    RETURN;                                    // 饱和即出口 / saturation is the exit
END_IF

// 段 8｜能力指数计算：六倍 σ 分母已由段 7 保证非零 / segment 8, capability indices
fSpan := DL_CPK_SIGMA_6 * fSigma;              // 双侧六倍标准差 / six sigma over both sides
fCp := (fUsl - fLsl) / fSpan;                  // 潜在能力 / potential capability
fUpper := (fUsl - fMean) / (DL_CPK_SIGMA_K * fSigma); // 上侧能力，分母同样过闸 / upper capability, the denominator passed the same gate
fLower := (fMean - fLsl) / (DL_CPK_SIGMA_K * fSigma); // 下侧能力 / lower capability
fCpk := MIN(fUpper, fLower);                   // 实际能力取两侧较小值 / actual capability takes the smaller side
fCp := MIN(fCp, fCpkSat);                      // 上侧饱和封顶 / cap the upside at the saturation limit
fCpk := MIN(fCpk, fCpkSat);                    // 上侧饱和封顶 / cap the upside at the saturation limit

// 段 9｜出口：返回 Cpk 并对位镜像 / segment 9, exit with the Cpk mirror
FC_DL_CpkIndex := fCpk;                        // 返回值即 Cpk / the return value is Cpk
bValid := TRUE;                                // 结果可用 / the result is usable
END_FUNCTION

(* ---- FC_DL_Crc16Generic.st ---- *)
(*
    组件名称 : FC_DL_Crc16Generic
    所属子库 : DL_MathData
    当前版本 : 1.0.1
    兼 容 性 : CODESYS V3.5+ / TwinCAT 3 / 汇川 InoProShop；仅依赖 Standard.library
    功能描述 : 参数化 CRC-16，poly / init / xorout / 输入反射 / 输出反射全部引脚化，一张实现覆盖任意从站协议。
              取舍 ①：参数化的动因 —— 库内 Crc16Modbus / Crc16Ccitt 把参数写死，遇到非标从站（自定义 poly 或只反射
              输入不反射输出）只能现场改源码，一改就失去可移植性；本件把参数域全部抬到引脚，算法内核只剩一份。
              取舍 ②：逐位算法，零查表零内存 —— 查表版快 8 倍但要 512 字节常量表，而跨平台移植时表初始化语法
              （数组常量初始化）恰恰是最容易踩坑的地方；本件优先可移植性，用 8 次定长位循环换「拷到任何平台都能编」。
              取舍 ③：反射不用专用位反指令 —— IEC 61131-3 没有标准位反函数，各平台扩展名不同；改用
              「右移 + 判最低位」的 8 次定长循环自建反射，只依赖 SHR/SHL/AND/OR。
              取舍 ④：帧长超上限拒绝而不截断 —— 截断后算出的 CRC 格式完全合法，却必然在校验端失败，
              这种「看起来对」的错误比明确报错贵得多。
    开源溯源 : T2-1 LGF CRC 子族，只借其参数域（initValue / finalXorValue / reflectInput / reflectResult）这一；本件为道莅 clean-room 防御性实现（仅借 LGF 分类事实/参数域/行为定义，零代码行与符号名复制）。
              分类级事实；逐位算法、反射实现、码位与错误分级 100% 自有，零代码行与注释复制。
    本文件内含 : FUNCTION FC_DL_Crc16Generic（单 POU，无配套类型）
    依 赖 : 无 DL_ 内部依赖；Standard.library: 无
    红线自检 : R1 ✓ 零全局变量与外部变量 ｜ R2 ✓ 零物理 IO 地址
              R3 ✓ 纯 IEC 61131-3 ｜ R4 ✓ 多项式零闸 + 帧长闸 + 空帧短路 + 位循环定长（无 WHILE、无需守卫）
              R5 ✓ 全变量中英双语同行注释 ｜ R6 N/A 纯函数无顺序状态机，无 CASE 可写
              R7 N/A 无定时器、无沿检测实例 ｜ R8 ✓ 位宽、循环边界、缓冲上限全常量化
    校验向量 : 对 ASCII "123456789"（9 字节，DL_CRC_VECT_LEN = 9）：
              ① CRC-16/ARC  poly=16#8005 init=16#0000 xorout=16#0000 入出双反射 → 16#BB3D
              ② CCITT-FALSE poly=16#1021 init=16#FFFF xorout=16#0000 不反射   → 16#29B1
              ③ XMODEM      poly=16#1021 init=16#0000 xorout=16#0000 不反射   → 16#31C3
              编码时以同构逐位算法做等价复算，三组向量全部命中（三元组与公开 CRC 参数目录一致）。
              任一不符即判定实现错误、禁止入库（R1 式规格向量错误防线）。
    错误码   : 16#0001_0445 [信息级] 空帧，返回 init XOR xorout，bValid = TRUE
               16#0001_0444 [信息级] 输出反射为真但多项式最高位为 0，疑似参数不匹配，bValid = TRUE
               16#0001_0384 [故障级] 多项式为零，CRC 无意义，返回 init XOR xorout，bValid = FALSE
               16#0001_0385 [故障级] 帧长超 DL_CRC_BUF_MAX，拒绝计算（不截断），返回 0，bValid = FALSE
               16#0001_0386 [故障级] 预留禁用（不得挪用）
    码位总账 : 16#0001_0445 用 / 16#0001_0444 用 ｜ 16#0001_0384 用 / 16#0001_0385 用 / 16#0001_0386 预留
    遗留假设 : ① 三组校验向量由等价算法脚本复算命中，未在 PLC 上实机运行 —— 属「算法已证、编译器未证」，
              交付门槛：须在 CODESYS / TwinCAT 3 / InoProShop 各编译并跑一次向量。
              ② WORD 上的 SHL/SHR 按 16 位容器截断（IEC 语义推导），若某平台按 32 位提升，位循环结果会偏离；
              该假设是本件唯一实质平台风险，需在门槛项里一并验证。
    修订历史 :
        2026-11-16  v1.0.0  首版，R21 批次 2 入库
        2026-11-16  v1.0.1  R21 终审修复（中等）：空帧分支原写 `uInit XOR uXorOut`，未过输出反射，
                            与本件自身的段 6 反射口径自相矛盾。零字节数据的正确结果应为
                            反射16(初值) XOR 终值：初值为回文（16#0000 / 16#FFFF）时两式同值，
                            非回文初值 + bReflectOut = TRUE 的参设下必错（典型如 init = 16#1234 的自定义从站）。
                            现空帧分支复用 16 次定长反射循环后再异或终值，与主体路径完全同构。
                            三组公开校验向量（非空帧）不受影响，仍为 BB3D / 29B1 / 31C3。
*)
FUNCTION FC_DL_Crc16Generic : WORD
VAR_INPUT
    nLen            : UINT;   // 待校验字节数，0~DL_CRC_BUF_MAX，0 = 空帧 [字节] / number of bytes, zero means an empty frame [byte]
    uPoly           : WORD;   // 生成多项式，如 16#8005 / 16#1021，为 0 即判故障 [无量纲] / generator polynomial, zero is a fault [dimensionless]
    uInit           : WORD;   // 寄存器初值 [无量纲] / initial register value [dimensionless]
    uXorOut         : WORD;   // 结果异或值 [无量纲] / final xor value [dimensionless]
    bReflectIn      : BOOL;   // 输入字节按位反射 / reflect every input byte
    bReflectOut     : BOOL;   // 结果 16 位反射 / reflect the sixteen bit result
END_VAR
VAR_IN_OUT
    afData          : ARRAY[0..DL_CRC_BUF_MAX] OF BYTE;   // 待校验字节数组，仅前 nLen 个有效 [字节] / data buffer, only the first nLen bytes are used [byte]
END_VAR
VAR_OUTPUT
    eErr            : UDINT;  // 错误码，0=正常；16#0001_04XX 信息级 / 16#0001_03XX 故障级 / error id, 0=ok
    bError          : BOOL;   // 故障级标志，eErr 落 16#0001_03XX 时为 TRUE / fault flag, TRUE on fault-level eErr
    bValid          : BOOL;   // 返回值是否可用 / result usable flag
END_VAR
VAR
    uCrc            : WORD;   // CRC 寄存器 [无量纲] / CRC register [dimensionless]
    uByte           : BYTE;   // 当前处理字节 [字节] / byte under processing [byte]
    uByteRefl       : WORD;   // 字节反射中间量 [位图] / byte reflection scratch [bitmap]
    uCrcRefl        : WORD;   // 结果反射中间量 [位图] / result reflection scratch [bitmap]
    uIdx            : UINT;   // 字节游标 [字节] / byte cursor [byte]
    nBit            : INT;    // 位游标 0~7 [位] / bit cursor 0..7 [bit]
    nReflBit        : INT;    // 反射循环位游标 0~15 [位] / reflection cursor 0..15 [bit]
END_VAR
VAR CONSTANT
    DL_CRC_BUF_MAX      : UINT := 255;                    // 单帧字节数上限（Modbus RTU / 645 远小于此）[字节] / frame length upper bound [byte]
    DL_CRC_BITS         : USINT := 16;                    // CRC 位宽，仅供上层核对位宽一致性；逻辑用 DL_CRC_REFL_LAST = 本值 − 1，故此处为说明性常量而非死码 [位] / CRC width kept as an advisory constant, the logic uses the last index instead [bit]
    DL_CRC_BIT_LAST     : INT := 7;                       // 字节位循环末值 [位] / last index of the byte bit loop [bit]
    DL_CRC_REFL_LAST    : INT := 15;                      // 结果反射循环末值 [位] / last index of the result reflection loop [bit]
    DL_CRC_SHIFT_BYTE   : INT := 8;                       // 字节左移量，恒为 8 [位] / constant left shift for one byte [bit]
    DL_CRC_LEN_NONE     : UINT := 0;                      // 空帧长度哨兵，减法前必判 [字节] / empty frame sentinel, tested before any subtraction [byte]
    DL_CRC_MSB_MASK     : WORD := 16#8000;                // 最高位掩码 [位图] / most significant bit mask [bitmap]
    DL_CRC_LSB_MASK     : WORD := 16#0001;                // 最低位掩码 [位图] / least significant bit mask [bitmap]
    DL_CRC_BYTE_MASK    : WORD := 16#00FF;                // 低字节掩码，反射结果收敛到字节 [位图] / low byte mask for the reflected byte [bitmap]
    DL_CRC_WORD_ZERO    : WORD := 16#0000;                // 零哨兵 [无量纲] / zero sentinel [dimensionless]
    DL_ERR_NONE         : UDINT := 16#0000_0000;          // 无故障 / no error
END_VAR

// 段 1｜返回值与错误状态预置 / segment 1, preset the return value and the error state
FC_DL_Crc16Generic := DL_CRC_WORD_ZERO;   // 故障缺省返回 0 / fault default returns zero
eErr   := DL_ERR_NONE;                    // 预置无错误 / preset no error
bError := FALSE;                          // 预置无故障 / preset no fault
bValid := FALSE;                          // 预置结果不可用 / preset unusable
uCrc   := uInit;                          // 寄存器装载初值 / load the initial value

// 段 2｜多项式闸：零多项式等于没有校验，必须拒算 / segment 2, zero polynomial gate
IF uPoly = DL_CRC_WORD_ZERO THEN
    FC_DL_Crc16Generic := uInit XOR uXorOut;   // 退化情形返回「初值异或终值」，口径与空帧一致 / degenerate case returns init xor xorout
    eErr   := 16#0001_0384;                    // 多项式为零（故障级）/ zero polynomial, fault level
    bError := TRUE;                            // 置故障标志 / raise the fault flag
    RETURN;                                    // bValid 保持 FALSE / bValid stays FALSE
END_IF

// 段 3｜帧长闸：超上限拒绝，绝不截断（截断的 CRC 必然校验失败却看着合法）/ segment 3, length gate, refuse instead of truncating
IF nLen > DL_CRC_BUF_MAX THEN
    FC_DL_Crc16Generic := DL_CRC_WORD_ZERO;    // 不给可疑结果 / never emit a suspicious result
    eErr   := 16#0001_0385;                    // 帧长超上限（故障级）/ frame too long, fault level
    bError := TRUE;                            // 置故障标志 / raise the fault flag
    RETURN;                                    // bValid 保持 FALSE / bValid stays FALSE
END_IF
IF nLen = DL_CRC_LEN_NONE THEN
    // 空帧同样必须过输出反射：寄存器一个字节都没进过，结果 = 反射16(初值) XOR 终值。
    // 漏这一步在初值为回文（16#0000 / 16#FFFF）时看不出差异，换非回文参设立刻错值，故不可省。
    uCrc := uInit;                             // 寄存器回到初值 / put the register back to the initial value
    IF bReflectOut THEN
        uCrcRefl := DL_CRC_WORD_ZERO;          // 反射累加器清零 / clear the reflection accumulator
        FOR nReflBit := 0 TO DL_CRC_REFL_LAST DO
            uCrcRefl := SHL(uCrcRefl, 1);                          // 左移腾位 / shift to make room
            uCrcRefl := uCrcRefl OR (uCrc AND DL_CRC_LSB_MASK);    // 取寄存器最低位 / take the lowest register bit
            uCrc     := SHR(uCrc, 1);                              // 寄存器右移 / shift the register down
        END_FOR
        uCrc := uCrcRefl;                      // 回写反射结果 / write the reflected value back
    END_IF
    FC_DL_Crc16Generic := uCrc XOR uXorOut;    // 空帧返回 反射(初值) XOR 终值（标准行为）/ an empty frame returns the reflected initial value xor xorout
    eErr   := 16#0001_0445;                    // 空帧（信息级，不置 bError）/ empty frame, info level
    bValid := TRUE;                            // 空帧是协议合法输入 / an empty frame is a legal protocol input
    RETURN;                                    // 提前出口，绝不进循环 / early exit, never enter the loop
END_IF

// 段 4｜反射参数一致性提示：输出反射却给了最高位为 0 的 poly，多半是参数抄错 / segment 4, reflection parameter sanity hint
IF bReflectOut AND ((uPoly AND DL_CRC_MSB_MASK) = DL_CRC_WORD_ZERO) THEN
    eErr := 16#0001_0444;                      // 反射参数与多项式最高位疑似不匹配（信息级）/ reflection parameter looks inconsistent, info level
END_IF

// 段 5｜逐字节位算法主体：nLen 已保证 ≥ 1，nLen − 1 不会回绕 / segment 5, byte by byte kernel, nLen is at least one
FOR uIdx := 0 TO nLen - 1 DO
    uByte := afData[uIdx];                     // 取当前字节，索引上界由长度闸保证 / fetch the byte, the upper bound is guaranteed by the length gate
    IF bReflectIn THEN
        uByteRefl := DL_CRC_WORD_ZERO;         // 反射累加器清零 / clear the reflection accumulator
        FOR nBit := 0 TO DL_CRC_BIT_LAST DO
            uByteRefl := SHL(uByteRefl, 1);                              // 左移腾位 / shift to make room
            uByteRefl := uByteRefl OR (BYTE_TO_WORD(uByte) AND DL_CRC_LSB_MASK);   // 取源字节最低位 / take the lowest source bit
            uByte     := SHR(uByte, 1);                                  // 源字节右移 / shift the source byte down
        END_FOR
        uByte := WORD_TO_BYTE(uByteRefl AND DL_CRC_BYTE_MASK);           // 收敛回一个字节 / converge back to one byte
    END_IF

    uCrc := uCrc XOR SHL(BYTE_TO_WORD(uByte), DL_CRC_SHIFT_BYTE);        // 字节置入高 8 位 / place the byte into the high half

    FOR nBit := 0 TO DL_CRC_BIT_LAST DO
        IF (uCrc AND DL_CRC_MSB_MASK) <> DL_CRC_WORD_ZERO THEN
            uCrc := SHL(uCrc, 1) XOR uPoly;    // 最高位为 1：左移后异或多项式 / top bit set, shift and xor the polynomial
        ELSE
            uCrc := SHL(uCrc, 1);              // 最高位为 0：只左移 / top bit clear, shift only
        END_IF
    END_FOR
END_FOR

// 段 6｜输出反射：16 次定长位循环，不用平台专用位反指令 / segment 6, output reflection with a fixed sixteen bit loop
IF bReflectOut THEN
    uCrcRefl := DL_CRC_WORD_ZERO;              // 反射累加器清零 / clear the reflection accumulator
    FOR nReflBit := 0 TO DL_CRC_REFL_LAST DO
        uCrcRefl := SHL(uCrcRefl, 1);                          // 左移腾位 / shift to make room
        uCrcRefl := uCrcRefl OR (uCrc AND DL_CRC_LSB_MASK);    // 取寄存器最低位 / take the lowest register bit
        uCrc     := SHR(uCrc, 1);                              // 寄存器右移 / shift the register down
    END_FOR
    uCrc := uCrcRefl;                          // 回写反射结果 / write the reflected value back
END_IF

// 段 7｜终值异或与出口 / segment 7, final xor and exit
FC_DL_Crc16Generic := uCrc XOR uXorOut;        // 异或终值 / apply the final xor
bValid := TRUE;                                // 结果可用 / the result is usable
END_FUNCTION

(* ---- FC_DL_Crc16Modbus.st ---- *)
(*==============================================================================
 * 组件名称 (Component)  : FC_DL_Crc16Modbus
 * 所属子库 (Sublibrary) : DL_MathData
 * 当前版本 (Version)    : 1.0.0
 * 兼容性   (Platform)   : CODESYS 3.5 / TwinCAT 3 / 汇川 InoProShop / Machine Expert
 *                         仅用标准 SHR / XOR / AND，无厂商方言、无查表常量数组
 * 功能描述 (Function)   : 标准 Modbus RTU CRC-16 校验计算。
 *                         参数：反射多项式 0xA001（即 0x8005 的位反转形式）、
 *                         初值 0xFFFF、输入输出反射（LSB first）、结果无异或。
 *                         逐位计算法：每字节先与 CRC 低字节异或，再循环 8 次
 *                         "取最低位 → 右移一位 → 若移出位为 1 则异或多项式"。
 *                         使用 SHR 而非除以 2，规避不同平台整数除法语义差异。
 * 算法     (Algorithm)  : 禁用除法取 LSB（B4），禁用点号位访问方言（B4），
 *                         必须先取最低位再右移（B5，顺序写反是最常见实现错误）。
 *
 * 【验收向量 / Acceptance vectors（已实算复核）】
 *   V1（本轮强制验收向量）
 *      帧  : 01 03 00 00 00 02
 *      CRC 寄存器值 = 16#0BC4，拼帧时按低字节先发：C4 0B
 *   V2  帧 01 03 00 00 00 0A  → 16#CDC5（发 C5 CD）
 *   V3  帧 11 03 00 6B 00 03  → 16#8776（发 76 87）
 *   V4  单字节 0x0C          → 16#45BF（发 BF 45）
 *
 * 【对 ROUND_PLAN §2.14 B7 的一处勘误 / Erratum】
 *   ROUND_PLAN 原文给出的单字节向量"0x0C → 0x911E"无法复现：按 Modbus 参数
 *   （初值 0xFFFF、反射多项式 0xA001）穷举 0..255 全部单字节输入，无任何取值
 *   得到 0x911E，故该值应源自其它多项式或其它初值的变体。本实现采用实算复核过的
 *   V4（0x0C → 0x45BF）替代，避免把错误向量写进单测造成"算法正确但测试失败"。
 *
 * 【返回字节序 / Byte order（B8）】
 *   函数返回的是 CRC 寄存器值（高字节在前语义）。拼帧时必须自行拆分：
 *     uCrc  := FC_DL_Crc16Modbus(abyData := aFrame, uByteCount := nLen);
 *     aFrame[nLen]     := WORD_TO_BYTE(uCrc AND 16#00FF);         「低字节先发」
 *     aFrame[nLen + 1] := WORD_TO_BYTE(SHR(uCrc, 8) AND 16#00FF); 「高字节后发」
 *
 * 【首版范围 / Scope of v1.0.0】
 *   仅实现逐位法，不含 256 项查表法：常量数组的跨平台初始化行为尚未验证，
 *   逐位法只有移位与异或两条语句，行为在三家平台上可预期。查表法列入 ROADMAP。
 * 开源溯源 (Origin)     : 原创实现。CRC-16/MODBUS 参数集见 Modbus over Serial Line
 *                         Specification V1.02 与公开 CRC 目录（Polynomial 0x8005 反射）。
 * 依赖     (Depends)    : 无 DL_ 内部依赖
 * 红线自检 (Redline)    : R1 ✓ 零全局变量表与外部变量引用 ｜ R2 ✓ 零物理 IO 地址直写
 *                         R3 ✓ 纯 IEC 61131-3（无除法取位、无点号位访问、显式 BYTE_TO_WORD）
 *                         R4 ✓ 长度为零/超限钳位 + 循环边界 + 位判断时序 + 下标校验
 *                         R5 ✓ 全变量中英双语同行注释 ｜ R6 N/A（无状态机）｜ R7 N/A（无实例调用）
 * 修订历史 (Revision)   :
 *   2026-11-14  v1.0.0  首版入库（Phase 1 冷启动 · Level 0 批次）
 *   2026-11-15  v1.0.1  R9 全库审计修复：头注释示例代码内嵌注释定界符改为引号形式，
 *                       消除"注释不可嵌套"平台上的提前闭合风险（算法与接口零变更）
 *============================================================================*)
FUNCTION FC_DL_Crc16Modbus : WORD
VAR_IN_OUT
    abyData : ARRAY[0..255] OF BYTE;   // 报文缓冲区，定长 256 字节，按 uByteCount 取前 N 字节 / Fixed 256-byte frame buffer, first N bytes are used
END_VAR
VAR_INPUT
    uByteCount : UINT := 0;            // 参与校验的字节数，合法域 1..256 / Number of bytes to checksum, valid range 1..256
END_VAR
VAR_OUTPUT
    bValid     : BOOL;                 // 长度合法标志，FALSE 表示已钳位或为零 / Length valid flag, FALSE means clamped or zero
    uErrorId   : UDINT;                // 故障码，0 = 无故障 / Error code, 0 = no error
END_VAR
VAR
    uCrc       : WORD;                 // CRC 寄存器，计算过程值 / CRC register, running value
    uCount     : UINT;                 // 钳位后的参与字节数 / Clamped byte count actually processed
    nIdx       : UINT;                 // 字节循环索引，值域 0..255 / Byte loop index, range 0..255
    nBit       : USINT;                // 位循环索引，固定 0..7 / Bit loop index, fixed 0..7
    bLsbSet    : BOOL;                 // 移位前最低位状态 / LSB state captured before the shift
END_VAR
VAR CONSTANT
    DL_CRC16_POLY   : WORD := 16#A001;   // 反射多项式 0x8005 / Reflected polynomial 0x8005
    DL_CRC16_INIT   : WORD := 16#FFFF;   // Modbus 规定初值 / Modbus mandated initial value
    DL_CRC16_MAXLEN : UINT := 256;       // 最大字节数，必须与数组维度一致 / Max byte count, must match the array dimension
END_VAR

(*------------------------------------------------------------------------------
 * 段 1｜安全预置：返回值先落到初值，异常路径下不得返回 0
 *      Safe preset: return falls back to the initial value, never to 0 on error paths
 *      0 在数学上是一个合法的 CRC 结果，返回它会让上层把"没算"误判成"算对了"
 *-----------------------------------------------------------------------------*)
FC_DL_Crc16Modbus := DL_CRC16_INIT;
bValid            := TRUE;
uErrorId          := 16#0000_0000;
uCrc              := DL_CRC16_INIT;
uCount            := uByteCount;

(*------------------------------------------------------------------------------
 * 段 2｜长度防御（边界 B1/B2）
 *      Length defence (boundaries B1/B2)
 *      零长度：返回初值 + 告警，直接退出（无字节可算）
 *      超限：钳到 256 后继续计算——现场排错时需要拿到一个可比对的值，
 *            中断会让诊断链断在第一步
 *-----------------------------------------------------------------------------*)
IF uByteCount = 0 THEN
    bValid   := FALSE;
    uErrorId := 16#0001_0001;
    RETURN;
ELSIF uByteCount > DL_CRC16_MAXLEN THEN
    uCount   := DL_CRC16_MAXLEN;
    bValid   := FALSE;
    uErrorId := 16#0001_0001;
END_IF

(*------------------------------------------------------------------------------
 * 段 3｜逐字节、逐位计算（边界 B3/B4/B5/B6）
 *      Byte-wise and bit-wise computation
 *      外层：uCount ≥ 1 已由段 2 保证，故 uCount - 1 不会下溢
 *      内层：固定 8 次，无动态步长、无 BY -1
 *      顺序硬约束：先取最低位 → 再右移 → 最后按标志异或
 *-----------------------------------------------------------------------------*)
FOR nIdx := 0 TO (uCount - 1) DO

    (* 数组下标上下界双检（红线 R4）：uCount ≤ 256 已保证 nIdx ≤ 255 *)
    (* Array index double check: uCount ≤ 256 guarantees nIdx ≤ 255 *)
    IF nIdx < DL_CRC16_MAXLEN THEN

        (* 显式 BYTE_TO_WORD 转换，禁止隐式提升（红线 R3） *)
        (* Explicit BYTE_TO_WORD conversion, implicit promotion is forbidden *)
        uCrc := uCrc XOR BYTE_TO_WORD(abyData[nIdx]);

        FOR nBit := 0 TO 7 DO
            (* 步骤 1：移位前先捕获最低位（边界 B5，顺序反了必然算错） *)
            (* Step 1: capture the LSB before shifting, reversing the order breaks the CRC *)
            bLsbSet := (uCrc AND 16#0001) <> 16#0000;

            (* 步骤 2：逻辑右移一位，禁用 / 2（边界 B4） *)
            (* Step 2: logical shift right by one, division by 2 is forbidden *)
            uCrc := SHR(uCrc, 1);

            (* 步骤 3：若移出位为 1，异或反射多项式 *)
            (* Step 3: if the shifted-out bit was 1, XOR the reflected polynomial *)
            IF bLsbSet THEN
                uCrc := uCrc XOR DL_CRC16_POLY;
            END_IF
        END_FOR;

    END_IF

END_FOR;

(*------------------------------------------------------------------------------
 * 段 4｜结果回写（边界 B8）：返回寄存器值，拆字节由调用方按低字节先发执行
 *      Result write-back: the register value is returned, byte splitting is the caller's job
 *-----------------------------------------------------------------------------*)
FC_DL_Crc16Modbus := uCrc;
END_FUNCTION

(* ---- FC_DL_Crc32Ethernet.st ---- *)
(*==============================================================================
 * 组件名称 (Component)  : FC_DL_Crc32Ethernet
 * 所属子库 (Sublibrary) : DL_MathData
 * 当前版本 (Version)    : 1.0.0
 * 兼容性   (Platform)   : CODESYS 3.5 / TwinCAT 3 / 汇川 InoProShop / Machine Expert
 *                         仅用标准 SHR / XOR / AND 与显式类型转换，无厂商方言
 * 功能描述 (Function)   : 标准 CRC-32/ISO-HDLC 校验码计算，即以太网 FCS、ZIP、PNG
 *                         使用的同一参数模型：反射多项式 16#EDB88320（即 16#04C11DB7
 *                         的位反射形式）、初值 16#FFFF_FFFF、终值异或 16#FFFF_FFFF。
 *                         逐位（bit-wise）实现：每字节先与 CRC 寄存器低 8 位异或，
 *                         再循环 8 次"取最低位 → 右移一位 → 移出位为 1 则异或多项式"。
 *                         支持分块链式调用：大报文分批计算，中间块 bFinalXor := FALSE，
 *                         把上一次返回值作为下一块的 uCrcSeed，最后一块才置 TRUE。
 *                         用于固件包完整性校验、文件传输校验、EtherCAT/Profinet 诊断
 *                         帧签核、上位机与 PLC 之间的报文校验。
 *
 * 【多项式方向警示 / Polynomial direction warning（边界 B1）】
 *   必须用反射值 16#EDB88320 配右移。若用 16#04C11DB7 配左移，得到的是
 *   CRC-32/BZIP2（"123456789" 算出 16#FC891918），两者不可混搭——
 *   混搭多项式方向是 CRC 实现的第一大错，且错误结果毫无规律可排查。
 *
 * 【链式调用契约 / Chained-call contract】
 *   分块时前 n-1 块传 bFinalXor := FALSE，把返回值直接作为下一块的 uCrcSeed；
 *   最后一块 bFinalXor := TRUE。中间块若误置 TRUE，相当于整体多异或了一次
 *   终值，整包校验必失败且极难定位（边界 B4）。
 *   调用序列文字说明（伪流程，非代码）：
 *     第 1 块：种子 = 默认全 1，末块标志 = FALSE，返回值记为 R1
 *     第 2 块：种子 = R1，末块标志 = FALSE，返回值记为 R2
 *     ……依此接力……
 *     第 n 块（末块）：种子 = R(n-1)，末块标志 = TRUE，返回值即整包 CRC
 *   分块大小可任意切分（含单字节），链式结果与一次性整包计算逐位一致。
 *
 * 【字节序披露 / Byte-order disclosure（边界 B7）】
 *   本函数只算数值。以太网 FCS 上帧时按小端（低字节先发）填入帧尾，
 *   拆字节与摆放顺序由组帧方决定，与本函数无关。
 *
 * 【扫描周期披露 / Cycle-time disclosure（边界 B5）】
 *   256 字节 × 8 位 = 2048 次内层循环，属重计算。应放在慢任务或事件触发
 *   任务中调用，不要放进 1 ms 高速任务拖垮总线周期。
 *
 * 【验收向量 / Acceptance vectors（已实算复核，算法独立交叉验证）】
 *   V1（本轮强制验收向量）
 *      "123456789"（31 32 33 34 35 36 37 38 39）
 *      seed 16#FFFF_FFFF、bFinalXor = TRUE → 16#CBF4_3926
 *   V2  空输入（nLength = 0）+ 默认参数 → 16#0000_0000（正确值，非错误）
 *   V3  单字节 00 → 16#D202_EF8D
 *   V4  分块链式："1234"（bFinalXor = FALSE，返回 16#641C_1F5C 作种子）
 *       + "56789"（bFinalXor = TRUE）→ 16#CBF4_3926（与 V1 一致，验证链式语义）
 *   V5  nLength = 300 → 钳位为 256 继续计算，nBytesUsed = 256，uErrorId = 16#0001_0001
 *
 * 【首版范围 / Scope of v1.0.0（边界 B6）】
 *   仅实现逐位法：零 RAM 开销、行为在三家平台可预期。若现场需要提速，
 *   按扩产规则另立 256 项查表变体，本组件内不加模式开关（禁止巨无霸）。
 * 开源溯源 (Origin)     : 依 IEEE 802.3 与公开 CRC 目录（CRC-32/ISO-HDLC 参数模型）
 *                         独立实现。OSCAT Network 校验函数族仅提供"按协议分族、
 *                         独立成函数"的组织方式参考（EPL-2.0）；其实现采用地址
 *                         指针入参，本库改为数组引脚传参，未复制任何源码。
 * 依赖     (Depends)    : 无 DL_ 内部依赖
 * 红线自检 (Redline)    : R1 ✓ 零全局变量表与外部变量引用 ｜ R2 ✓ 零物理 IO 地址直写
 *                         R3 ✓ 纯 IEC 61131-3（显式 BYTE_TO_DWORD，无位访问方言）
 *                         R4 ✓ 长度钳位 + 下标双检 + 空输入兜底（空输入是合法值）
 *                         R5 ✓ 全变量中英双语同行注释 ｜ R6 N/A（无状态机）｜ R7 N/A（无实例调用）
 * 修订历史 (Revision)   :
 *   2026-11-14  v1.0.0  首版入库（Phase 1 收口批次 · R3）
 *============================================================================*)
FUNCTION FC_DL_Crc32Ethernet : DWORD
VAR_IN_OUT
    aabyData   : ARRAY[0..255] OF BYTE;   // 待校验字节缓冲，定长 256，按 nLength 取前 N 字节 / Fixed 256-byte data buffer, first nLength bytes are used
END_VAR
VAR_INPUT
    nLength    : INT;                     // 本次参与计算的字节数，合法域 0..256，越界自动钳位 / Byte count this call, range 0..256, clamped
    uCrcSeed   : DWORD := 16#FFFF_FFFF;   // 初值或上一分块的返回值（链式调用），首块用默认值 / Initial value or previous chunk result for chaining
    bFinalXor  : BOOL  := TRUE;           // TRUE = 输出前异或 16#FFFF_FFFF，仅最后一块置 TRUE / Final XOR, TRUE on the last chunk only
END_VAR
VAR_OUTPUT
    uErrorId   : UDINT;                   // 故障码，0 = 无故障，16#0001_0001 = 长度越界已钳位 / Error code, 0 = no error, 0001_0001 = length clamped
    nBytesUsed : INT;                     // 实际参与计算的字节数（钳位后），供诊断 / Bytes actually processed after clamping
END_VAR
VAR
    uCrc       : DWORD;                   // CRC 工作寄存器 / CRC working register
    nLenWork   : INT;                     // 钳位后的本地长度副本，不回写输入引脚 / Local clamped copy of the length
    nI         : INT;                     // 字节循环索引，值域 0..255 / Byte loop index, range 0..255
    nBit       : INT;                     // 位循环索引，固定 8 次 / Bit loop index, fixed 8 iterations
    uByte      : DWORD;                   // 当前字节零扩展到 32 位 / Current byte zero-extended to 32 bits
    bLsbSet    : BOOL;                    // 右移前最低位状态 / LSB state captured before the shift
END_VAR
VAR CONSTANT
    DL_CRC32_POLY_REFLECTED : DWORD := 16#EDB8_8320;  // IEEE 802.3 多项式 16#04C11DB7 的位反射形式 / Bit-reflected IEEE 802.3 polynomial
    DL_CRC32_INIT           : DWORD := 16#FFFF_FFFF;  // 参数模型规定初值，全 1 / Mandated all-ones initial value
    DL_CRC32_XOROUT         : DWORD := 16#FFFF_FFFF;  // 终值异或值 / Final XOR value
    DL_CRC32_BUF_MAX        : INT   := 256;           // 缓冲上限，必须与数组维度一致 / Buffer limit, must match the array dimension
    DL_CRC32_BITS_PER_BYTE  : INT   := 8;             // 每字节位循环次数 / Bit iterations per byte
    DL_CRC32_BIT_MASK       : DWORD := 16#0000_0001;  // 最低位提取掩码 / LSB extraction mask
END_VAR

(*------------------------------------------------------------------------------
 * 段 1｜安全预置：返回值先落初值，故障码清零，长度取本地副本
 *      Safe preset: return value falls back to the seed, error code cleared
 *-----------------------------------------------------------------------------*)
FC_DL_Crc32Ethernet := uCrcSeed;
uErrorId            := 16#0000_0000;
nBytesUsed          := 0;
uCrc                := uCrcSeed;
nLenWork            := nLength;

(*------------------------------------------------------------------------------
 * 段 2｜长度防御（边界 B3/B5）：钳位而非拒绝，让诊断链拿到可比对的值
 *      Length defence: clamp instead of reject so diagnostics still get a value
 *      负值 → 0；大于 256 → 256；均置 16#0001_0001（瞬时码）
 *-----------------------------------------------------------------------------*)
IF nLenWork < 0 THEN
    nLenWork := 0;
    uErrorId := 16#0001_0001;
ELSIF nLenWork > DL_CRC32_BUF_MAX THEN
    nLenWork := DL_CRC32_BUF_MAX;
    uErrorId := 16#0001_0001;
END_IF

(*------------------------------------------------------------------------------
 * 段 3｜逐字节、逐位计算（边界 B1）
 *      Byte-wise and bit-wise computation
 *      顺序硬约束：先与寄存器低 8 位异或 → 循环 8 次
 *      （先捕获最低位 → 右移 → 移出位为 1 则异或反射多项式）
 *      空输入（nLenWork = 0）跳过循环，返回值为终值异或后的 16#0000_0000，
 *      这是参数模型的正确结果而非错误（边界 B3）
 *-----------------------------------------------------------------------------*)
IF nLenWork > 0 THEN

    FOR nI := 0 TO (nLenWork - 1) DO

        (* 数组下标上下界双检（红线 R4）：nLenWork ≤ 256 已保证 nI ≤ 255 *)
        (* Array index double check: nLenWork ≤ 256 guarantees nI ≤ 255 *)
        IF nI < DL_CRC32_BUF_MAX THEN

            (* 显式 BYTE_TO_DWORD 零扩展，禁止隐式提升（红线 R3） *)
            (* Explicit BYTE_TO_DWORD zero extension, implicit promotion is forbidden *)
            uByte := BYTE_TO_DWORD(aabyData[nI]);
            uCrc  := uCrc XOR uByte;

            FOR nBit := 1 TO DL_CRC32_BITS_PER_BYTE DO
                (* 步骤 1：右移前先捕获最低位，顺序反了必然算错 *)
                (* Step 1: capture the LSB before shifting, reversing breaks the CRC *)
                bLsbSet := (uCrc AND DL_CRC32_BIT_MASK) <> 16#0000_0000;

                (* 步骤 2：逻辑右移一位，禁用除法取位（红线 R3） *)
                (* Step 2: logical shift right by one, division is forbidden *)
                uCrc := SHR(uCrc, 1);

                (* 步骤 3：若移出位为 1，异或反射多项式 *)
                (* Step 3: if the shifted-out bit was 1, XOR the reflected polynomial *)
                IF bLsbSet THEN
                    uCrc := uCrc XOR DL_CRC32_POLY_REFLECTED;
                END_IF
            END_FOR;

        END_IF

    END_FOR;

END_IF

(*------------------------------------------------------------------------------
 * 段 4｜终值与回写：仅最后一块做终值异或（链式契约见头注释）
 *      Final value and write-back: final XOR only on the last chunk
 *-----------------------------------------------------------------------------*)
IF bFinalXor THEN
    uCrc := uCrc XOR DL_CRC32_XOROUT;
END_IF

nBytesUsed          := nLenWork;
FC_DL_Crc32Ethernet := uCrc;

(*------------------------------------------------------------------------------
 * 段 5｜自检断言说明（供单元测试与现场对拍，向量已实算复核）
 *      Self-check assertion notes for unit tests and on-site cross-checks
 *      V1  "123456789"，种子默认、末块标志 TRUE → 16#CBF4_3926
 *      V2  空输入（长度 0），种子默认、末块标志 TRUE → 16#0000_0000
 *      V3  单字节 00，种子默认、末块标志 TRUE → 16#D202_EF8D
 *      V4  "1234"（末块标志 FALSE，返回 16#641C_1F5C 作种子）
 *          + "56789"（末块标志 TRUE）→ 16#CBF4_3926，与 V1 逐位一致
 *      V5  长度传 300 → 钳位为 256 继续计算，本函数输出 16#0001_0001
 *          且 nBytesUsed = 256，返回值为前 256 字节的校验值
 *-----------------------------------------------------------------------------*)
END_FUNCTION
